(* IEC 61131-3 sources: PLC-IsaVODE/PLC-IsaVODE/samples/plc-programs (part 2) *)

(* ---- 251-SETUP_LANGUAGE.ST ---- *)
TYPE oscat_LANGUAGE:
	STRUCT
		DEFAULT 	: INT;
		LMAX    	: INT;
	END_STRUCT;
END_TYPE

FUNCTION_BLOCK SETUP_LANGUAGE_Block

	VAR_IN_OUT
		LANGUAGE :	oscat_LANGUAGE;
	END_VAR

	VAR
		init :	BOOL;
	END_VAR

	IF init THEN RETURN; END_IF;
	init := TRUE;

	LANGUAGE.DEFAULT  := 1; (* 1=english, 2=german 3=french *)
	LANGUAGE.LMAX := 3;

END_FUNCTION_BLOCK

PROGRAM program0

	VAR
		LANGUAGE :	oscat_LANGUAGE;
		func_block : SETUP_LANGUAGE_Block;
	END_VAR
		func_block.LANGUAGE  := LANGUAGE;
		func_block();
		LANGUAGE := func_block.LANGUAGE;

END_PROGRAM

CONFIGURATION Config0

	RESOURCE Res0 ON PLC
		TASK task0(INTERVAL := T#20ms,PRIORITY := 0);
		PROGRAM instance0 WITH task0 : program0;
	END_RESOURCE

END_CONFIGURATION

(* ---- 253-ENERGY.ST ---- *)
FUNCTION_BLOCK ENERGY
	VAR_INPUT
		J :	REAL;
		C :	REAL;
		WH :	REAL;
	END_VAR

	VAR_OUTPUT
		YJ :	REAL;
		YC :	REAL;
		YWH :	REAL;
	END_VAR

	YJ := J + Wh * 3600.0 + C * 4.1868;
	YC := YJ * 0.238845896627496;
	YWh := YJ * 2.7777777778E-004;
END_FUNCTION_BLOCK

PROGRAM program0
  VAR
		J  :	REAL;
		C  :	REAL;
		WH :	REAL;

		YJ  :	REAL;
		YC  :	REAL;
		YWH :	REAL;
	func_block : ENERGY;
  END_VAR
	func_block.J  :=J ;
	func_block.C  :=C ;
	func_block.WH :=WH;
	func_block();
	YJ  := func_block.YJ ;
	YC  := func_block.YC ;
	YWH := func_block.YWH;

END_PROGRAM

CONFIGURATION Config0
	RESOURCE Res0 ON PLC
		TASK task0(INTERVAL := T#20ms,PRIORITY := 0);
		PROGRAM instance0 WITH task0 : program0;
	END_RESOURCE
END_CONFIGURATION

(* ---- 257-FINDB_NONUM.ST ---- *)
FUNCTION_BLOCK FINDB_NONUM_Block

	VAR_INPUT
		STR :	STRING;
	END_VAR

	VAR_OUTPUT
		FINDB_NONUM :	INT;
	END_VAR

	VAR
		pos :	INT;
		x :	INT;
	END_VAR

	pos := LEN(str);
	WHILE (pos >=1) DO
		x :=GET_CHAR(str,pos);
		IF (X < 48 AND X <> 46) OR X > 57 THEN
			findB_nonum := pos;
			RETURN;
		END_IF;
	pos := pos -1;
	END_WHILE;
	findB_nonum := 0;

END_FUNCTION_BLOCK

PROGRAM program0
	VAR
		STR :	STRING;

		FINDB_NONUM :	INT;

		func_block : FINDB_NONUM_Block;
	END_VAR
	func_block.STR := STR;
	func_block();
	FINDB_NONUM  := func_block.FINDB_NONUM;
END_PROGRAM

CONFIGURATION Config0
	RESOURCE Res0 ON PLC
		TASK task0(INTERVAL := T#20ms,PRIORITY := 0);
		PROGRAM instance0 WITH task0 : program0;
	END_RESOURCE
END_CONFIGURATION

(* ---- 258-HYST_1.ST ---- *)
FUNCTION_BLOCK HYST_1_Block

	VAR_INPUT
		IN :	REAL;
		HIGH :	REAL;
		LOW :	REAL;
	END_VAR

	VAR_OUTPUT
		Q :	BOOL;
		WIN :	BOOL;
	END_VAR

	IF in < low THEN
		Q := FALSE;
		win := FALSE;
	ELSIF in > high THEN
		Q := TRUE;
		win := FALSE;
	ELSE
		win := TRUE;
	END_IF;

END_FUNCTION_BLOCK

PROGRAM program0
	VAR
		IN :	REAL;
		HIGH :	REAL;
		LOW :	REAL;
		Q :	BOOL;
		WIN :	BOOL;
		func_block : HYST_1_Block;
	END_VAR
	func_block.IN := IN;
	func_block.HIGH := HIGH;
	func_block.LOW := LOW;
	func_block();
	Q  := func_block.Q;
	WIN  := func_block.WIN;
END_PROGRAM

CONFIGURATION Config0
	RESOURCE Res0 ON PLC
		TASK task0(INTERVAL := T#20ms,PRIORITY := 0);
		PROGRAM instance0 WITH task0 : program0;
	END_RESOURCE
END_CONFIGURATION

(* ---- 260-V3_SUB.ST ---- *)
TYPE oscat_vector_3:
	STRUCT
		X : REAL;
		Y : REAL;
		Z : REAL;
	END_STRUCT;
END_TYPE

FUNCTION_BLOCK V3_SUB_Block

	VAR_INPUT
		A :	oscat_vector_3;
		B :	oscat_vector_3;
	END_VAR

	VAR_OUTPUT
		V3_SUB :	oscat_vector_3;
	END_VAR

	V3_SUB.X := A.X - B.X;
	V3_SUB.Y := A.Y - B.Y;
	V3_SUB.Z := A.Z - B.Z;

END_FUNCTION_BLOCK

PROGRAM program0
  	VAR
		A :	oscat_vector_3;
		B :	oscat_vector_3;
		V3_SUB :	oscat_vector_3;
		func_block : V3_SUB_Block;
  	END_VAR
	func_block.A := A;
	func_block.B := B;
	func_block();
	V3_SUB := func_block.V3_SUB;
END_PROGRAM

CONFIGURATION Config0
  RESOURCE Res0 ON PLC
    TASK task0(INTERVAL := T#20ms,PRIORITY := 0);
    PROGRAM instance0 WITH task0 : program0;
  END_RESOURCE
END_CONFIGURATION

(* ---- 261-A_TRIG.ST ---- *)
FUNCTION_BLOCK A_TRIG

	VAR_INPUT
		IN :	REAL;
		RES :	REAL;
	END_VAR

	VAR_OUTPUT
		Q :	BOOL;
		D :	REAL;
	END_VAR

	VAR
		last_in :	REAL;
	END_VAR

	D := IN - LAST_IN;
	IF ABS(D) >= res THEN
		Q := TRUE;
		last_in := IN;
	ELSE
		Q := FALSE;
	END_IF;

END_FUNCTION_BLOCK

PROGRAM program0
	VAR
	    LocalVar0 : REAL;
		LocalVar1 : REAL;
		LocalOUT1  : BOOL;
		LocalOUT2  : REAL;
		func_block : A_TRIG;
  	END_VAR
	func_block.IN := LocalVar0;
    func_block.RES := LocalVar1;
	func_block();
	LocalOUT1 := func_block.Q;
	LocalOUT2 := func_block.D;
END_PROGRAM

CONFIGURATION Config0
  	RESOURCE Res0 ON PLC
    	TASK task0(INTERVAL := T#20ms,PRIORITY := 0);
    	PROGRAM instance0 WITH task0 : program0;
  	END_RESOURCE
END_CONFIGURATION

(* ---- 265-INTERLOCK.ST ---- *)
FUNCTION_BLOCK INTERLOCK_Block

	VAR_INPUT
		I1 :	BOOL;
		I2 :	BOOL;
		TL :	TIME;
	END_VAR

	VAR_OUTPUT
		Q1 :	BOOL;
		Q2 :	BOOL;
	END_VAR

	VAR
		T1 :	TOF;
		T2 :	TOF;
	END_VAR

	T1(IN := I1, PT := TL);
	T2(IN := I2, PT := TL);

	Q1 := I1 AND NOT t2.Q;
	Q2 := I2 AND NOT t1.Q;

END_FUNCTION_BLOCK

PROGRAM program0
	VAR
		I1 :	BOOL;
		I2 :	BOOL;
		TL :	TIME;
		Q1 :	BOOL;
		Q2 :	BOOL;
		func_block : INTERLOCK_Block;
  	END_VAR
	func_block.I1  :=I1;
	func_block.I2  :=I2;
	func_block.TL  :=TL;
	func_block();
	Q1 := func_block.Q1;
	Q2 := func_block.Q2;
END_PROGRAM

CONFIGURATION Config0
	RESOURCE Res0 ON PLC
		TASK task0(INTERVAL := T#20ms,PRIORITY := 0);
		PROGRAM instance0 WITH task0 : program0;
	END_RESOURCE
END_CONFIGURATION

(* ---- 266-CMUL.ST ---- *)
TYPE oscat_complex :
  STRUCT
	re : REAL;
	im : REAL;
  END_STRUCT;
END_TYPE

FUNCTION_BLOCK CMUL_Block

	VAR_INPUT
		X :	oscat_complex;
		Y :	oscat_complex;
	END_VAR

	VAR_OUTPUT
		CMUL :	oscat_complex;
	END_VAR

	CMUL.re := X.re * Y.re - X.im * Y.im;
	CMUL.im := X.re * Y.im + X.im * Y.re;
END_FUNCTION_BLOCK

PROGRAM program0
  VAR
    LocalVar0 : oscat_complex;
	LocalVar1 : oscat_complex;
	LocalOUT  : oscat_complex;
	func_block : CMUL_Block;
  END_VAR
	func_block.X  := LocalVar0;
	func_block.Y  := LocalVar1;
	func_block();
	LocalOUT := func_block.CMUL;
END_PROGRAM

CONFIGURATION Config0
  RESOURCE Res0 ON PLC
    TASK task0(INTERVAL := T#20ms,PRIORITY := 0);
    PROGRAM instance0 WITH task0 : program0;
  END_RESOURCE
END_CONFIGURATION

(* ---- 268-IS_UPPER.ST ---- *)
FUNCTION SETUP_EXTENDED_ASCII:BOOL

	VAR_INPUT
		X :	BOOL;
	END_VAR

	SETUP_EXTENDED_ASCII := X OR TRUE;

END_FUNCTION

FUNCTION ISC_UPPER:BOOL

	VAR_INPUT
		IN :	BYTE;
	END_VAR

	IF SETUP_EXTENDED_ASCII(FALSE) THEN
		ISC_UPPER :=  ((in > BYTE#64) AND (in < BYTE#91)) OR (((in > BYTE#191) AND (in < BYTE#223)) AND (in <> BYTE#215));
	ELSE
		ISC_UPPER := ((in > BYTE#64) AND (in < BYTE#91));
	END_IF;

END_FUNCTION

FUNCTION_BLOCK IS_UPPER

	VAR_INPUT
		STR :	STRING;
	END_VAR

	VAR_OUTPUT
		IS_UPPER :	BOOL;
	END_VAR

	VAR
		pos :	INT;
		I :	INT;
	END_VAR

	I := LEN(str);
	FOR pos := 1 TO I DO
		IF NOT ISC_UPPER(INT_TO_BYTE(GET_CHAR(str,pos))) THEN
			IS_UPPER := FALSE;
			RETURN;
		END_IF;
	END_FOR;
	IS_UPPER := I>0;

END_FUNCTION_BLOCK

(* ---- 269-IS_CC.ST ---- *)
FUNCTION_BLOCK IS_CC_Block

	VAR_INPUT
		STR :	STRING;
		CMP :	STRING;
	END_VAR

	VAR_OUTPUT
		IS_CC :	BOOL;
	END_VAR

	VAR
		L :	INT;
		pos :	INT;
		temp :	STRING;
	END_VAR

	L := LEN(str);
	FOR pos := 1 TO L DO
		temp := MID(str,1,pos);
		IF FIND(CMP,temp) = 0 THEN
			IS_CC := FALSE;
			RETURN;
		END_IF;
	END_FOR;
	IS_CC := L > 0;

END_FUNCTION_BLOCK

PROGRAM program0

	VAR
		STR :	STRING;
		CMP :	STRING;

		IS_CC :	BOOL;

		func_block : IS_CC_Block;
	END_VAR
	func_block.STR := STR;
	func_block.CMP := CMP;
	func_block();
	IS_CC := func_block.IS_CC;

END_PROGRAM

CONFIGURATION Config0

	RESOURCE Res0 ON PLC
		TASK task0(INTERVAL := T#20ms,PRIORITY := 0);
		PROGRAM instance0 WITH task0 : program0;
	END_RESOURCE

END_CONFIGURATION

(* ---- 271-IS_NCC.ST ---- *)
FUNCTION_BLOCK IS_NCC_Block

	VAR_INPUT
		STR :	STRING;
		CMP :	STRING;
	END_VAR

	VAR_OUTPUT
		IS_NCC :	BOOL;
	END_VAR

	VAR
		L :	INT;
		pos :	INT;
		temp :	STRING;
	END_VAR

	L := LEN(str);
	FOR pos := 1 TO L DO
		temp := MID(str,1,pos);
		IF FIND(CMP,temp) > 0 THEN
			IS_NCC := FALSE;
			RETURN;
		END_IF;
	END_FOR;
	IS_NCC := TRUE;

END_FUNCTION_BLOCK

PROGRAM program0

	VAR
		STR :	STRING;
		CMP :	STRING;
		IS_NCC :	BOOL;
		func_block : IS_NCC_Block;
	END_VAR
	func_block.STR := STR;
	func_block.CMP := CMP;
	func_block();
	IS_NCC := func_block.IS_NCC;

END_PROGRAM

CONFIGURATION Config0

	RESOURCE Res0 ON PLC
		TASK task0(INTERVAL := T#20ms,PRIORITY := 0);
		PROGRAM instance0 WITH task0 : program0;
	END_RESOURCE

END_CONFIGURATION

(* ---- 273-TONOF.ST ---- *)
FUNCTION_BLOCK TONOF

	VAR_INPUT
		IN :	BOOL;
		T_ON :	TIME;
		T_OFF :	TIME;
	END_VAR

	VAR_OUTPUT
		Q :	BOOL;
	END_VAR

	VAR
		X :	TON;
		old :	BOOL;
		mode :	BOOL;
	END_VAR

	IF IN XOR old THEN
	X(IN := FALSE, PT := SEL_TIME(IN,T_OFF,T_ON));
	mode := IN;
	old := IN;
	END_IF;
	X(IN := TRUE);
	IF X.Q THEN Q := mode;END_IF;

END_FUNCTION_BLOCK

PROGRAM program0
  VAR
	IN :	BOOL;
	T_ON :	TIME;
	T_OFF :	TIME;
	Q :	BOOL;
	func_block : TONOF;
  END_VAR
	func_block.IN  :=IN ;
	func_block.T_ON  :=T_ON ;
	func_block.T_OFF  :=T_OFF ;
	func_block();
	Q := func_block.Q;

END_PROGRAM

CONFIGURATION Config0
	RESOURCE Res0 ON PLC
		TASK task0(INTERVAL := T#20ms,PRIORITY := 0);
		PROGRAM instance0 WITH task0 : program0;
	END_RESOURCE
END_CONFIGURATION

(* ---- 278-DWORD_TO_STRB.ST ---- *)
FUNCTION_BLOCK DWORD_TO_STRB_Block
	VAR_INPUT
		IN :	DWORD;
	END_VAR

	VAR_OUTPUT
		DWORD_TO_STRB :	STRING;
	END_VAR

	VAR
		i :	INT;
	END_VAR

	DWORD_TO_STRB :='';
	FOR i := 1 TO 32 DO
		IF (in AND DWORD#16#8000_0000) > DWORD#0 THEN
			DWORD_TO_STRB := CONCAT(DWORD_TO_STRB,'1');
		ELSE
			DWORD_TO_STRB := CONCAT(DWORD_TO_STRB,'0');
		END_IF;
		in := SHL(in, 1);
	END_FOR;
END_FUNCTION_BLOCK

PROGRAM program0
  VAR
    IN :	DWORD;

	DWORD_TO_STRB :	STRING;
	func_block : DWORD_TO_STRB_Block;
  END_VAR
	func_block.IN  := IN;
	func_block();
	DWORD_TO_STRB := func_block.DWORD_TO_STRB;
END_PROGRAM

CONFIGURATION Config0
  RESOURCE Res0 ON PLC
    TASK task0(INTERVAL := T#20ms,PRIORITY := 0);
    PROGRAM instance0 WITH task0 : program0;
  END_RESOURCE
END_CONFIGURATION

(* ---- 279-STAIR2.ST ---- *)
FUNCTION FLOOR : INT
	VAR_INPUT
		x : REAL;
	END_VAR

	FLOOR := REAL_TO_INT(X);
	IF INT_TO_REAL(FLOOR) > X THEN
		floor := floor - 1;
	END_IF;
END_FUNCTION

FUNCTION_BLOCK STAIR2_Block

	VAR_INPUT
		X :	REAL;
		D :	REAL;
	END_VAR

	VAR_OUTPUT
		Y :	REAL;
	END_VAR

	IF D > 0.0 THEN
		IF X >= Y + D OR X <= Y - D THEN Y := INT_TO_REAL(FLOOR(X/D)) * D; END_IF;
	ELSE
		Y := X;
	END_IF;

END_FUNCTION_BLOCK

PROGRAM program0

	VAR
		X :	REAL;
		D :	REAL;
		Y :	REAL;
		func_block : STAIR2_Block;
	END_VAR
	func_block.X := X;
	func_block.D := D;
	func_block();
	Y := func_block.Y;

END_PROGRAM

CONFIGURATION Config0

	RESOURCE Res0 ON PLC
		TASK task0(INTERVAL := T#20ms,PRIORITY := 0);
		PROGRAM instance0 WITH task0 : program0;
	END_RESOURCE

END_CONFIGURATION

(* ---- 280-DEC_TO_BYTE.ST ---- *)
FUNCTION_BLOCK DEC_TO_BYTE_Block
	VAR_INPUT
		DEC :	STRING;
	END_VAR

	VAR_OUTPUT
		DEC_TO_BYTE :	BYTE;
	END_VAR

	VAR
		i :	INT;
		X :	INT;
		stop :	INT;
	END_VAR

	DEC_TO_BYTE := BYTE#0;
	stop := LEN(DEC);
	FOR I := 1 TO stop DO
		X := GET_CHAR(DEC,I);
		IF X > 47 AND X < 58 THEN
			DEC_TO_BYTE := INT_TO_BYTE(_BYTE_TO_INT(DEC_TO_BYTE) * 10 + X - 48);
		END_IF;
	END_FOR;

END_FUNCTION_BLOCK

PROGRAM program0
  VAR
    LocalVar0 : STRING;
	LocalOUT  : BYTE;
	func_block : DEC_TO_BYTE_Block;
  END_VAR
	func_block.DEC  := LocalVar0;
	func_block();
	LocalOUT := func_block.DEC_TO_BYTE;
END_PROGRAM

CONFIGURATION Config0
  RESOURCE Res0 ON PLC
    TASK task0(INTERVAL := T#20ms,PRIORITY := 0);
    PROGRAM instance0 WITH task0 : program0;
  END_RESOURCE
END_CONFIGURATION

(* ---- 281-BYTE_TO_STRB.ST ---- *)
FUNCTION_BLOCK BYTE_TO_STRB_Block
	VAR_INPUT
		IN :	BYTE;
	END_VAR

	VAR_OUTPUT
		BYTE_TO_STRB :	STRING;
	END_VAR

	VAR
		i :	INT;
	END_VAR

	BYTE_TO_STRB := '';
	FOR i := 1 TO 8 DO
		IF (in AND BYTE#2#1000_0000) = BYTE#2#1000_0000 THEN
			BYTE_TO_STRB := CONCAT(BYTE_TO_STRB,'1');
		ELSE
			BYTE_TO_STRB := CONCAT(BYTE_TO_STRB,'0');
		END_IF;
		in := SHL(in, 1);
	END_FOR;

END_FUNCTION_BLOCK

PROGRAM program0
  VAR
    LocalVar0 : BYTE;
	LocalOUT  : STRING;
	func_block : BYTE_TO_STRB_Block;
  END_VAR
	func_block.IN  := LocalVar0;
	func_block();
	LocalOUT := func_block.BYTE_TO_STRB;

END_PROGRAM

CONFIGURATION Config0
  RESOURCE Res0 ON PLC
    TASK task0(INTERVAL := T#20ms,PRIORITY := 0);
    PROGRAM instance0 WITH task0 : program0;
  END_RESOURCE
END_CONFIGURATION

(* ---- 282-SW_RECONFIG.ST ---- *)
FUNCTION_BLOCK SW_RECONFIG_Block

	VAR_INPUT
		IN :	BOOL;
		TD :	TIME;
		TR :	TIME;
	END_VAR

	VAR_OUTPUT
		Q :	BOOL;
	END_VAR

	VAR
		T1 :	TON;
		T2 :	TON;
		INV :	BOOL;
	END_VAR

	t1(in := IN, PT := TD);

	IF tr > t#0s THEN
		Q := t1.Q XOR inv;
		T2(in := Q, pt := TR);
		IF T2.Q THEN INV := NOT INV; END_IF;
	ELSE
		Q := t1.Q;
	END_IF;

END_FUNCTION_BLOCK

PROGRAM program0
	VAR
		IN :	BOOL;
		TD :	TIME;
		TR :	TIME;
		Q :	BOOL;

		func_block : SW_RECONFIG_Block;
	END_VAR
	func_block.IN := IN;
	func_block.TD := TD;
	func_block.TR := TR ;

	func_block();
	Q  := func_block.Q;

END_PROGRAM

CONFIGURATION Config0
	RESOURCE Res0 ON PLC
		TASK task0(INTERVAL := T#20ms,PRIORITY := 0);
		PROGRAM instance0 WITH task0 : program0;
	END_RESOURCE
END_CONFIGURATION

(* ---- 283-CINV.ST ---- *)
TYPE oscat_complex :
  STRUCT
	re : REAL;
	im : REAL;
  END_STRUCT;
END_TYPE

FUNCTION_BLOCK CINV_Block

	VAR_INPUT
		X :	oscat_complex;
	END_VAR

	VAR_OUTPUT
		CINV :	oscat_complex;
	END_VAR

	VAR
		temp :	REAL;
	END_VAR

	temp := X.re * X.re + X.im * X.im;
	IF temp = 0.0 THEN CINV.re := 0.0;CINV.im := 0.0;RETURN;END_IF;
	CINV.re := X.re / temp;
	CINV.im := -X.im / temp;

END_FUNCTION_BLOCK

PROGRAM program0
  VAR
    LocalVar0 : oscat_complex;
	LocalOUT  : oscat_complex;
	func_block : CINV_Block;
  END_VAR
	func_block.X  := LocalVar0;
	func_block();
	LocalOUT := func_block.CINV;
END_PROGRAM

CONFIGURATION Config0
  RESOURCE Res0 ON PLC
    TASK task0(INTERVAL := T#20ms,PRIORITY := 0);
    PROGRAM instance0 WITH task0 : program0;
  END_RESOURCE
END_CONFIGURATION

(* ---- 284-V3_XPRO.ST ---- *)
TYPE oscat_vector_3 :
	STRUCT
		X : REAL;
		Y : REAL;
		Z : REAL;
	END_STRUCT;
END_TYPE

FUNCTION_BLOCK V3_XPRO_Block
	VAR_INPUT
		A :	oscat_vector_3;
		B :	oscat_vector_3;
	END_VAR

	VAR_OUTPUT
		V3_XPRO :	oscat_vector_3;
	END_VAR

	V3_XPRO.X := A.Y * B.Z - A.Z * B.Y;
	V3_XPRO.Y := A.Z * B.X - A.X * B.Z;
	V3_XPRO.Z := A.X * B.Y - A.Y * B.X;

END_FUNCTION_BLOCK

PROGRAM program0
  	VAR
		A :	oscat_vector_3;
		B :	oscat_vector_3;
		V3_XPRO :	oscat_vector_3;
		func_block : V3_XPRO_Block;
  	END_VAR
	func_block.A := A;
	func_block.B := B;
	func_block();
	V3_XPRO := func_block.V3_XPRO;
END_PROGRAM

CONFIGURATION Config0
  RESOURCE Res0 ON PLC
    TASK task0(INTERVAL := T#20ms,PRIORITY := 0);
    PROGRAM instance0 WITH task0 : program0;
  END_RESOURCE
END_CONFIGURATION

(* ---- 288-DEC_4.ST ---- *)
FUNCTION_BLOCK DEC_4
	VAR_INPUT
		D :	BOOL;
		A0 :	BOOL;
		A1 :	BOOL;
	END_VAR

	VAR_OUTPUT
		Q0 :	BOOL;
		Q1 :	BOOL;
		Q2 :	BOOL;
		Q3 :	BOOL;
	END_VAR

	Q0 := D AND NOT A0 AND NOT A1;
	Q1 := D AND A0 AND NOT A1;
	Q2 := D AND NOT A0 AND A1;
	Q3 := D AND A0 AND A1;
END_FUNCTION_BLOCK

PROGRAM program0
  VAR
	D :	BOOL;
	A0 :	BOOL;
	A1 :	BOOL;

	Q0 :	BOOL;
	Q1 :	BOOL;
	Q2 :	BOOL;
	Q3 :	BOOL;

	func_block : DEC_4;
  END_VAR
	func_block.D   := D  ;
	func_block.A0  := A0  ;
	func_block.A1  := A1  ;
	func_block();
	Q0:= func_block.Q0;
	Q1:= func_block.Q1;
	Q2:= func_block.Q2;
	Q3:= func_block.Q3;
END_PROGRAM

CONFIGURATION Config0
  RESOURCE Res0 ON PLC
    TASK task0(INTERVAL := T#20ms,PRIORITY := 0);
    PROGRAM instance0 WITH task0 : program0;
  END_RESOURCE
END_CONFIGURATION

(* ---- 291-FF_D2E.ST ---- *)
FUNCTION_BLOCK FF_D2E
	VAR_INPUT
		D0 :	BOOL;
		D1 :	BOOL;
		CLK :	BOOL;
		RST :	BOOL;
	END_VAR

	VAR_OUTPUT
		Q0 :	BOOL;
		Q1 :	BOOL;
	END_VAR

	VAR
		edge :	BOOL;
	END_VAR

	IF rst THEN
		Q0 := FALSE;
		Q1 := FALSE;
	ELSIF clk AND NOT edge THEN
		Q0 := D0;
		Q1 := D1;
	END_IF;
	edge := CLK;

END_FUNCTION_BLOCK

PROGRAM program0
  VAR
	D0  :	BOOL;
	D1  :	BOOL;
	CLK :	BOOL;
	RST :	BOOL;

	Q0 :	BOOL;
	Q1 :	BOOL;

	func_block : FF_D2E;
  END_VAR
	func_block.D0  :=D0 ;
	func_block.D1  :=D1 ;
	func_block.CLK :=CLK;
	func_block.RST :=RST;
	func_block();
	Q0 := func_block.Q0;
	Q1 := func_block.Q1;
END_PROGRAM

CONFIGURATION Config0
  RESOURCE Res0 ON PLC
    TASK task0(INTERVAL := T#20ms,PRIORITY := 0);
    PROGRAM instance0 WITH task0 : program0;
  END_RESOURCE
END_CONFIGURATION

(* ---- 292-HYST_2.ST ---- *)
FUNCTION_BLOCK HYST_2_Block

	VAR_INPUT
		IN :	REAL;
		VAL :	REAL;
		HYS :	REAL;
	END_VAR

	VAR_OUTPUT
		Q :	BOOL;
		WIN :	BOOL;
	END_VAR

	VAR
		tmp :	REAL;
	END_VAR

	tmp := val - hys * 0.5;
	IF in < tmp THEN
		Q := FALSE;
		win := FALSE;
	ELSIF in > tmp + hys THEN
		Q := TRUE;
		win := FALSE;
	ELSE
		win := TRUE;
	END_IF;

END_FUNCTION_BLOCK

PROGRAM program0
	VAR
		IN :	REAL;
		VAL :	REAL;
		HYS :	REAL;
		Q :	BOOL;
		WIN :	BOOL;
		func_block : HYST_2_Block;
	END_VAR
	func_block.IN := IN;
	func_block.VAL := VAL;
	func_block.HYS := HYS;
	func_block();
	Q  := func_block.Q;
	WIN  := func_block.WIN;
END_PROGRAM

CONFIGURATION Config0
	RESOURCE Res0 ON PLC
		TASK task0(INTERVAL := T#20ms,PRIORITY := 0);
		PROGRAM instance0 WITH task0 : program0;
	END_RESOURCE
END_CONFIGURATION

(* ---- 294-FF_RSE.ST ---- *)
FUNCTION_BLOCK FF_RSE
	VAR_INPUT
		CS :	BOOL;
		CR :	BOOL;
		RST :	BOOL;
	END_VAR

	VAR_OUTPUT
		Q :	BOOL;
	END_VAR

	VAR
		es :	BOOL;
		er :	BOOL;
	END_VAR

	IF rst THEN
		(* asynchronous reset *)
		Q := FALSE;
	ELSIF CR AND NOT er THEN
		(* rising edge on CR *)
		Q := FALSE;
	ELSIF CS AND NOT es THEN
		(* rising edge on CS *)
		Q := TRUE;
	END_IF;

	es := CS;
	er := CR;
END_FUNCTION_BLOCK

PROGRAM program0
  VAR
	CS  :	BOOL;
	CR  :	BOOL;
	RST :	BOOL;

	Q :	BOOL;

	func_block : FF_RSE;
  END_VAR
	func_block.CS  :=CS ;
	func_block.CR  :=CR ;
	func_block.RST :=RST;
	func_block();
	Q := func_block.Q;
END_PROGRAM

CONFIGURATION Config0
  RESOURCE Res0 ON PLC
    TASK task0(INTERVAL := T#20ms,PRIORITY := 0);
    PROGRAM instance0 WITH task0 : program0;
  END_RESOURCE
END_CONFIGURATION

(* ---- 296-BUFFER_CLEAR_NW.ST ---- *)
TYPE
  oscat_NW_BUF_LONG  : ARRAY [0..4095] OF BYTE;
END_TYPE

FUNCTION_BLOCK _BUFFER_CLEAR_NW
	VAR_INPUT
		SIZE :	UINT;
	END_VAR

	VAR_OUTPUT
		BUFFER_CLEAR :	BOOL;
	END_VAR

	VAR_IN_OUT
		PT :	oscat_NW_BUF_LONG;
	END_VAR

	VAR
		err :	INT;
		result :	WORD;
	END_VAR
	result:=MEMSET(err,BYTE#00,UINT_TO_DINT(size),pt[0]);
	BUFFER_CLEAR := (err = 0);
END_FUNCTION_BLOCK

PROGRAM program0
  VAR
	SIZE :	UINT;

	BUFFER_CLEAR :	BOOL;

	PT :	oscat_NW_BUF_LONG;

	func_block : _BUFFER_CLEAR_NW;
  END_VAR
	func_block.SIZE  :=SIZE ;
	func_block.PT  :=PT ;
	func_block();
	PT := func_block.PT;
	BUFFER_CLEAR := func_block.BUFFER_CLEAR;
END_PROGRAM

CONFIGURATION Config0
  RESOURCE Res0 ON PLC
    TASK task0(INTERVAL := T#20ms,PRIORITY := 0);
    PROGRAM instance0 WITH task0 : program0;
  END_RESOURCE
END_CONFIGURATION

(* ---- 298-FF_JKE.ST ---- *)
FUNCTION_BLOCK FF_JKE
	VAR_INPUT
		SET :	BOOL;
		J :	BOOL;
		CLK :	BOOL;
		K :	BOOL;
		RST :	BOOL;
	END_VAR

	VAR_OUTPUT
		Q :	BOOL;
	END_VAR

	VAR
		edge :	BOOL;
	END_VAR

	IF rst OR set THEN
		Q := NOT rst;
	ELSIF clk AND NOT edge THEN
		IF J XOR K THEN Q := J;
		ELSE Q := K XOR Q;
		END_IF;
	END_IF;
	edge := CLK;

END_FUNCTION_BLOCK

PROGRAM program0
  VAR
		SET :	BOOL;
		J   :	BOOL;
		CLK :	BOOL;
		K   :	BOOL;
		RST :	BOOL;

		Q :	BOOL;

	func_block : FF_JKE;
  END_VAR
	func_block.SET :=SET;
	func_block.J   :=J  ;
	func_block.CLK :=CLK;
	func_block.K   :=K  ;
	func_block.RST :=RST;
	func_block();
	Q := func_block.Q;
END_PROGRAM

CONFIGURATION Config0
  RESOURCE Res0 ON PLC
    TASK task0(INTERVAL := T#20ms,PRIORITY := 0);
    PROGRAM instance0 WITH task0 : program0;
  END_RESOURCE
END_CONFIGURATION

(* ---- 299-OCT_TO_DWORD.ST ---- *)
FUNCTION_BLOCK OCT_TO_DWORD_Block

	VAR_INPUT
		OCT :	STRING;
	END_VAR

	VAR_OUTPUT
		OCT_TO_DWORD :	DWORD;
	END_VAR

	VAR
		i :	INT;
		stop :	INT;
		X :	INT;
	END_VAR

	OCT_TO_DWORD := DWORD#0;
	stop := LEN(oct);
	FOR I := 1 TO stop DO
		X := GET_CHAR(oct,I);
		(* calculate the value of the digit *)
		IF X > 47 AND x < 56 THEN
			OCT_TO_DWORD := SHL_DWORD(OCT_TO_DWORD,3) OR INT_TO_DWORD(X - 48);
		END_IF;
	END_FOR;

END_FUNCTION_BLOCK

PROGRAM program0
  VAR
    OCT : STRING;
    OCT_TO_DWORD : DWORD;
	func_block : OCT_TO_DWORD_Block;
  END_VAR

  	func_block.OCT := '125';
	func_block();
	OCT_TO_DWORD := func_block.OCT_TO_DWORD;
END_PROGRAM

CONFIGURATION Config0
	RESOURCE Res0 ON PLC
		TASK task0(INTERVAL := T#20ms,PRIORITY := 0);
		PROGRAM instance0 WITH task0 : program0;
	END_RESOURCE
END_CONFIGURATION

(* ---- 3-IS_LOWER.ST ---- *)
FUNCTION_BLOCK IS_LOWER

VAR_INPUT
	STR :	STRING;
END_VAR

VAR_OUTPUT
	IS_LOWER :	BOOL;
END_VAR

VAR
	pos :	INT;
	I :	INT;
END_VAR

I := LEN(str);
FOR pos := 1 TO I DO
	IF NOT ISC_LOWER(INT_TO_BYTE(GET_CHAR(str,pos))) THEN
		IS_LOWER := FALSE;
		RETURN;
	END_IF;
END_FOR;
IS_LOWER := I>0;

END_FUNCTION_BLOCK

(* ---- 302-MD5_TO_STRH.ST ---- *)
FUNCTION_BLOCK MD5_TO_STRH

	VAR_INPUT
		MD5 :	oscat_aB0_15;
	END_VAR

	VAR_OUTPUT
		MD5_TO_STRH :	oscat_STRING32;
	END_VAR

	VAR
		buf :	oscat_aB0_31;
		x :	INT;
		BUF_TO_STRING :	BUF_TO_STRING;
		i :	INT;
		tmp :	INT;
	END_VAR

	x := 0;
	FOR i := 0 TO 15 DO;
		tmp := BYTE_TO_INT(SHR_BYTE(MD5[i],4));
		buf[x] := INT_TO_BYTE(tmp + SEL(tmp <= 9,87,48));
		x := x + 1;
		tmp := BYTE_TO_INT(MD5[i] AND BYTE#2#1111);
		buf[x] := INT_TO_BYTE(tmp + SEL(tmp <= 9,87,48));
		x := x + 1;
	END_FOR;

	FOR x := 0 TO 1 DO
		BUF_TO_STRING.REQ := x > 0;
		BUF_TO_STRING.BUF_FORMAT := TRUE;
		BUF_TO_STRING.BUF_OFFS := DINT#0;
		BUF_TO_STRING.BUF_CNT := DINT#32;
		BUF_TO_STRING.BUFFER := buf;
		BUF_TO_STRING.DST := MD5_TO_STRH;
		BUF_TO_STRING();
		buf := BUF_TO_STRING.BUFFER;
		MD5_TO_STRH := BUF_TO_STRING.DST;
	END_FOR;

END_FUNCTION_BLOCK

(* ---- 303-FINDB.ST ---- *)
FUNCTION_BLOCK FINDB_Block

	VAR_INPUT
		STR1 :	STRING;
		STR2 :	STRING;
	END_VAR

	VAR_OUTPUT
		FINDB :	INT;
	END_VAR

	VAR
		pos :	INT;
		length :	INT;
		string_temp :	STRING;
	END_VAR

	length := LEN(str2);
	pos := LEN(str1) - length +1;
	WHILE (pos >= 1) DO
		string_temp := MID(str1,length,pos);
		IF EQ_STRING(string_temp,str2) THEN
			FindB := pos;
			RETURN;
		END_IF;
	pos := pos -1;
	END_WHILE;
	FindB := 0;

END_FUNCTION_BLOCK

PROGRAM program0
  VAR
		STR1 :	STRING;
		STR2 :	STRING;

		FINDB :	INT;

	func_block : FINDB_Block;
  END_VAR
	func_block.STR1  := STR1;
	func_block.STR2  := STR2;
	func_block();
	FINDB := func_block.FINDB;
END_PROGRAM

CONFIGURATION Config0

	RESOURCE Res0 ON PLC
		TASK task0(INTERVAL := T#20ms,PRIORITY := 0);
		PROGRAM instance0 WITH task0 : program0;
	END_RESOURCE
END_CONFIGURATION

(* ---- 305-SEL2_OF_3B.ST ---- *)
FUNCTION_BLOCK SEL2_OF_3B_Block

	VAR_INPUT
		IN1 :	BOOL;
		IN2 :	BOOL;
		IN3 :	BOOL;
		TD :	TIME;
	END_VAR

	VAR_OUTPUT
		Q :	BOOL;
		W :	BOOL;
	END_VAR

	VAR
		TDEL :	TON;
	END_VAR

	Q := (IN1 AND IN2) OR (IN1 AND IN3) OR (IN2 AND IN3);
	TDEL(IN := (in1 XOR in2) OR (in1 XOR in3) OR (in2 XOR in3), PT := TD);
	W := TDEL.Q;

END_FUNCTION_BLOCK

PROGRAM program0

	VAR
		IN1 :	BOOL;
		IN2 :	BOOL;
		IN3 :	BOOL;
		TD :	TIME;
		Q :	BOOL;
		W :	BOOL;
		func_block : SEL2_OF_3B_Block;
  	END_VAR
	func_block.IN1  :=IN1;
	func_block.IN2  :=IN2;
	func_block.IN3  :=IN3;
	func_block.TD  :=TD;
	func_block();
	Q := func_block.Q;
	W := func_block.W;

END_PROGRAM

CONFIGURATION Config0

	RESOURCE Res0 ON PLC
		TASK task0(INTERVAL := T#20ms,PRIORITY := 0);
		PROGRAM instance0 WITH task0 : program0;
	END_RESOURCE

END_CONFIGURATION

(* ---- 306-ARRAY_SUM.ST ---- *)
TYPE
	oscat_pt_ARRAY: ARRAY [1..100] OF REAL;
END_TYPE

FUNCTION_BLOCK ARRAY_SUM_Block
	VAR_IN_OUT
		PT :	oscat_pt_ARRAY;
	END_VAR

	VAR_INPUT
		SIZE :	UINT;
	END_VAR

	VAR_OUTPUT
		ARRAY_SUM :	REAL;
	END_VAR

	VAR
		i :	INT;
		stop :	INT;
	END_VAR

	stop :=LIMIT_INT(1,UINT_TO_INT(size),1000);

	array_sum := pt[1];
	FOR i := 2 TO stop DO
		array_sum := array_sum + pt[i];
	END_FOR;
END_FUNCTION_BLOCK

PROGRAM program0
  VAR
    LocalVar0 : oscat_pt_ARRAY;
    LocalVar1 : UINT;
	LocalOUT  : REAL;
	func_block : ARRAY_SUM_Block;
  END_VAR
	func_block.pt := LocalVar0;
	func_block.size := LocalVar1;
	func_block();
	LocalOUT := func_block.ARRAY_SUM;

END_PROGRAM

CONFIGURATION Config0
  RESOURCE Res0 ON PLC
    TASK task0(INTERVAL := T#20ms,PRIORITY := 0);
    PROGRAM instance0 WITH task0 : program0;
  END_RESOURCE
END_CONFIGURATION

(* ---- 307-ARRAY_MAX.ST ---- *)
TYPE
	oscat_pt_ARRAY: ARRAY [1..100] OF REAL;
END_TYPE

FUNCTION_BLOCK ARRAY_MAX_Block
	VAR_IN_OUT
		PT :	oscat_pt_ARRAY;
	END_VAR

	VAR_INPUT
		SIZE :	UINT;
	END_VAR

	VAR_OUTPUT
		ARRAY_MAX :	REAL;
	END_VAR

	VAR
		i :	INT;
		stop :	INT;
	END_VAR

	stop :=LIMIT_INT(1,UINT_TO_INT(size),1000);

	FOR i := 1 TO stop DO
		IF pt[i] > array_max THEN array_max := pt[i]; END_IF;
	END_FOR;

END_FUNCTION_BLOCK

PROGRAM program0
  VAR
    LocalVar0 : oscat_pt_ARRAY;
    LocalVar1 : UINT;
	LocalOUT  : REAL;
	func_block : ARRAY_MAX_Block;
  END_VAR
	func_block.pt := LocalVar0;
	func_block.size := LocalVar1;
	func_block();
	LocalOUT := func_block.ARRAY_MAX;

END_PROGRAM

CONFIGURATION Config0
  RESOURCE Res0 ON PLC
    TASK task0(INTERVAL := T#20ms,PRIORITY := 0);
    PROGRAM instance0 WITH task0 : program0;
  END_RESOURCE
END_CONFIGURATION

(* ---- 308-DWORD_TO_STRF.ST ---- *)
FUNCTION_BLOCK DWORD_TO_STRF_Block

	VAR_INPUT
		IN :	DWORD;
		N :	INT;
	END_VAR

	VAR_OUTPUT
		DWORD_TO_STRF :	STRING;
	END_VAR

	VAR
		temp :	STRING;
		temp2 :	STRING;
		L : INT;
	END_VAR

	temp := DWORD_TO_STRING(in);
	L := LEN(temp);
	IF N < L THEN
		temp :=RIGHT(temp,N);
		L := N;
	END_IF;

	WHILE L < N DO
		temp2 := temp;
		temp := CONCAT('0', temp2);
		L := L + 1;
	END_WHILE;
	DWORD_TO_STRF := temp;

END_FUNCTION_BLOCK

PROGRAM program0
  VAR
    IN :	DWORD;
	N :		INT;
	DWORD_TO_STRF :	STRING;
	func_block : DWORD_TO_STRF_Block;
  END_VAR
	func_block.IN  := IN;
	func_block.N  := N;
	func_block();
	DWORD_TO_STRF := func_block.DWORD_TO_STRF;
END_PROGRAM

CONFIGURATION Config0
  RESOURCE Res0 ON PLC
    TASK task0(INTERVAL := T#20ms,PRIORITY := 0);
    PROGRAM instance0 WITH task0 : program0;
  END_RESOURCE
END_CONFIGURATION

(* ---- 309-SHA1_TO_STRH.ST ---- *)
FUNCTION_BLOCK SHA1_TO_STRH_Block

	VAR_INPUT
		SHA1 :	oscat_aB0_19;
	END_VAR

	VAR_OUTPUT
		SHA1_TO_STRH :	oscat_STRING40;
	END_VAR

	VAR
		buf :	oscat_aB0_39;
		i :	INT;
		tmp :	INT;
		x :	INT;
		BUF_TO_STRING :	BUF_TO_STRING;
	END_VAR

	x := 0;
	FOR i := 0 TO 19 DO;
		tmp := BYTE_TO_INT(SHR_BYTE(SHA1[i],4));
		buf[x] := INT_TO_BYTE(tmp + SEL(tmp <= 9,87,48));
		x := x + 1;
		tmp := BYTE_TO_INT(SHA1[i] AND BYTE#2#1111);
		buf[x] := INT_TO_BYTE(tmp + SEL(tmp <= 9,87,48));
		x := x + 1;
	END_FOR;

	FOR x := 0 TO 1 DO
		BUF_TO_STRING.REQ := x > 0;
		BUF_TO_STRING.BUF_FORMAT := TRUE;
		BUF_TO_STRING.BUF_OFFS := DINT#0;
		BUF_TO_STRING.BUF_CNT := DINT#40;
		BUF_TO_STRING.BUFFER := buf;
		BUF_TO_STRING.DST := SHA1_TO_STRH;
		BUF_TO_STRING();
		buf := BUF_TO_STRING.BUFFER;
		SHA1_TO_STRH := BUF_TO_STRING.DST;
	END_FOR;

END_FUNCTION_BLOCK

(* ---- 311-CLEAN.ST ---- *)
FUNCTION_BLOCK CLEAN_Block
	VAR_INPUT
		IN :	STRING;
		CX :	STRING;
	END_VAR

	VAR_OUTPUT
		CLEAN :	STRING;
	END_VAR

	VAR
		pos :	INT;
		stop :	INT;
		char :	STRING;
	END_VAR

	CLEAN := IN;
	stop := LEN(in);
	pos := 1;
	WHILE pos <= stop DO
		char := MID(CLEAN, 1, pos);
		IF FIND(cx,char) > 0 THEN
			pos := pos + 1;
		ELSE
			CLEAN := DELETE(CLEAN, 1, pos);
			stop := stop - 1;
		END_IF;
	END_WHILE;

END_FUNCTION_BLOCK

PROGRAM program0
  VAR
    LocalVar0 : STRING;
    LocalVar1 : STRING;
	LocalOUT  : STRING;
	func_block : CLEAN_Block;
  END_VAR
	func_block.IN  := LocalVar0;
	func_block.CX := LocalVar1;
	func_block();
	LocalOUT := func_block.CLEAN;

END_PROGRAM

CONFIGURATION Config0
  RESOURCE Res0 ON PLC
    TASK task0(INTERVAL := T#20ms,PRIORITY := 0);
    PROGRAM instance0 WITH task0 : program0;
  END_RESOURCE
END_CONFIGURATION

(* ---- 312-COUNT_SUBSTRING.ST ---- *)
FUNCTION_BLOCK COUNT_SUBSTRING_Block
	VAR_INPUT
		SEARCH :	STRING;
		STR :	STRING;
	END_VAR

	VAR_OUTPUT
		COUNT_SUBSTRING :	INT;
	END_VAR

	VAR
		pos :	INT;
		size :	INT;
	END_VAR

	COUNT_SUBSTRING := 0;
	size := LEN(SEARCH);
	REPEAT
	pos := FIND(STR,SEARCH);
	IF pos > 0 THEN
		STR := REPLACE(STR, '', size,pos);
		COUNT_SUBSTRING := COUNT_SUBSTRING + 1;
	END_IF;
	UNTIL pos = 0
	END_REPEAT;
END_FUNCTION_BLOCK

PROGRAM program0
  VAR
	SEARCH :	STRING;
	STR :	STRING;

	COUNT_SUBSTRING :	INT;
	func_block : COUNT_SUBSTRING_Block;
  END_VAR
	func_block.SEARCH  :=SEARCH  ;
	func_block.STR   :=STR   ;

	func_block();
	COUNT_SUBSTRING := func_block.COUNT_SUBSTRING;
END_PROGRAM

CONFIGURATION Config0
  RESOURCE Res0 ON PLC
    TASK task0(INTERVAL := T#20ms,PRIORITY := 0);
    PROGRAM instance0 WITH task0 : program0;
  END_RESOURCE
END_CONFIGURATION

(* ---- 313-CDIV.ST ---- *)
TYPE oscat_complex :
  STRUCT
	re : REAL;
	im : REAL;
  END_STRUCT;
END_TYPE

FUNCTION_BLOCK CDIV_Block

	VAR_INPUT
		X :	oscat_complex;
		Y :	oscat_complex;
	END_VAR

	VAR_OUTPUT
		CDIV :	oscat_complex;
	END_VAR

	VAR
		temp :	REAL;
	END_VAR

	temp := Y.re * Y.re + Y.im * Y.im;
	IF temp = 0.0 THEN CDIV.re := 0.0;CDIV.im := 0.0;RETURN;END_IF;
	CDIV.re := (X.re * Y.re + X.im * Y.im) / temp;
	CDIV.im := (X.im * Y.re - X.re * Y.im) / temp;

END_FUNCTION_BLOCK

PROGRAM program0

	VAR
		X :	oscat_complex;
		Y :	oscat_complex;

		CDIV :	oscat_complex;

		func_block : CDIV_Block;
	END_VAR
	func_block.X := X;
	func_block.Y := Y;
	func_block();
	CDIV := func_block.CDIV;

END_PROGRAM

CONFIGURATION Config0

	RESOURCE Res0 ON PLC
		TASK task0(INTERVAL := T#20ms,PRIORITY := 0);
		PROGRAM instance0 WITH task0 : program0;
	END_RESOURCE

END_CONFIGURATION

(* ---- 314-TO_UML.ST ---- *)
FUNCTION _BYTE_TO_INT:INT
	VAR_INPUT
		IN :	BYTE;
	END_VAR

	_BYTE_TO_INT := USINT_TO_INT(BYTE_TO_USINT(IN));
END_FUNCTION

FUNCTION_BLOCK TO_UML_Block

	VAR_INPUT
		IN :	BYTE;
	END_VAR

	VAR_OUTPUT
		TO_UML :	STRING;
	END_VAR

	CASE _BYTE_TO_INT(in) OF
		196:
			TO_UML := 'Ae';
		214:
			TO_UML := 'Oe';
		220:
			TO_UML := 'Ue';
		223:
			TO_UML := 'ss';
		228:
			TO_UML := 'ae';
		246:
			TO_UML := 'oe';
		252:
			TO_UML := 'ue';
	ELSE
		TO_UML := BYTE_TO_STRING(IN);
	END_CASE;

END_FUNCTION_BLOCK

PROGRAM program0
  VAR
	IN :	BYTE;
	TO_UML :	STRING;
	func_block : TO_UML_Block;
  END_VAR
	func_block.IN  := IN;
	func_block();
	TO_UML := func_block.TO_UML;

END_PROGRAM

CONFIGURATION Config0
	RESOURCE Res0 ON PLC
		TASK task0(INTERVAL := T#20ms,PRIORITY := 0);
		PROGRAM instance0 WITH task0 : program0;
	END_RESOURCE
END_CONFIGURATION

(* ---- 315-ARRAY_MIN.ST ---- *)
TYPE
	oscat_pt_ARRAY: ARRAY [1..100] OF REAL;
END_TYPE

FUNCTION_BLOCK ARRAY_MIN_Block
	VAR_IN_OUT
		PT :	oscat_pt_ARRAY;
	END_VAR

	VAR_INPUT
		SIZE :	UINT;
	END_VAR

	VAR_OUTPUT
		ARRAY_MIN :	REAL;
	END_VAR

	VAR
		i :	INT;
		stop :	INT;
	END_VAR

	stop :=LIMIT_INT(1,UINT_TO_INT(size),1000);

	array_min := pt[1];
	FOR i := 2 TO stop DO
		IF pt[i] < array_min THEN array_min := pt[i]; END_IF;
	END_FOR;

END_FUNCTION_BLOCK
PROGRAM program0
  VAR
    LocalVar0 : oscat_pt_ARRAY;
    LocalVar1 : UINT;
	LocalOUT  : REAL;
	func_block : ARRAY_MIN_Block;
  END_VAR
	func_block.pt := LocalVar0;
	func_block.size := LocalVar1;
	func_block();
	LocalOUT := func_block.ARRAY_MIN;

END_PROGRAM

CONFIGURATION Config0
  RESOURCE Res0 ON PLC
    TASK task0(INTERVAL := T#20ms,PRIORITY := 0);
    PROGRAM instance0 WITH task0 : program0;
  END_RESOURCE
END_CONFIGURATION

(* ---- 316-LOWERCASE.ST ---- *)
FUNCTION_BLOCK LOWERCASE_Block

	VAR_INPUT
		STR :	STRING;
	END_VAR

	VAR_OUTPUT
		LOWERCASE :	STRING;
	END_VAR

	VAR
		char :	BYTE;
		char2 :	BYTE;
		pos :	INT;
		l :	INT;
		str_temp :	STRING;
	END_VAR

	LOWERCASE := str;
	l := LEN(str);
	FOR pos := 1 TO l DO
		char := INT_TO_BYTE(GET_CHAR(str,pos));
		char2 := TO_LOWER(char);
		IF char <> char2 THEN
			str_temp := LOWERCASE;
			LOWERCASE := REPLACE(str_temp,BYTE_TO_STRING(char2,'%c'),1,pos);
		END_IF;
	END_FOR;

END_FUNCTION_BLOCK

PROGRAM program0
  VAR
    OCT : STRING;
    LOWERCASE : STRING;
	func_block : LOWERCASE_Block;
  END_VAR

  	func_block.OCT := '125';
	func_block();
	LOWERCASE := func_block.LOWERCASE;
END_PROGRAM

CONFIGURATION Config0
	RESOURCE Res0 ON PLC
		TASK task0(INTERVAL := T#20ms,PRIORITY := 0);
		PROGRAM instance0 WITH task0 : program0;
	END_RESOURCE
END_CONFIGURATION

(* ---- 318-UPPERCASE.ST ---- *)
FUNCTION_BLOCK UPPERCASE_Block

	VAR_INPUT
		STR :	STRING;
	END_VAR

	VAR_OUTPUT
		UPPERCASE :	STRING;
	END_VAR

	VAR
		char :	BYTE;
		char2 :	BYTE;
		pos :	INT;
		l :	INT;
		str_temp :	STRING;
	END_VAR

	UPPERCASE := str;
	l := LEN(str);
	FOR pos := 1 TO l DO
		char := INT_TO_BYTE(GET_CHAR(str,pos));
		char2 := TO_UPPER(char);
		IF char <> char2 THEN
			str_temp := UPPERCASE;
			UPPERCASE := REPLACE(str_temp,BYTE_TO_STRING(char2,'%c'),1,pos);
		END_IF;
	END_FOR;

END_FUNCTION_BLOCK

PROGRAM program0
	VAR
	    LocalVar1 : STRING;
		LocalOUT  : STRING;
		func_block : UPPERCASE_Block;
  	END_VAR
	func_block.STR := LocalVar1;
	func_block();
	LocalOUT := func_block.UPPERCASE;
END_PROGRAM

CONFIGURATION Config0
  	RESOURCE Res0 ON PLC
    	TASK task0(INTERVAL := T#20ms,PRIORITY := 0);
    	PROGRAM instance0 WITH task0 : program0;
  	END_RESOURCE
END_CONFIGURATION

(* ---- 319-CLICK_CNT.ST ---- *)
FUNCTION_BLOCK CLICK_CNT
	VAR_INPUT
		IN :	BOOL;
		N :	INT;
		TC :	TIME;
	END_VAR

	VAR_OUTPUT
		Q :	BOOL;
	END_VAR

	VAR
		tx :	TP;
		edge :	BOOL;
		cnt :	INT := INT#-1;
	END_VAR

	Q := FALSE;

	IF in AND NOT edge AND NOT tx.q THEN
		cnt := 0;
	ELSIF tx.Q AND NOT IN AND edge THEN
		cnt := cnt + 1;
	ELSIF NOT tx.Q THEN
		Q := cnt=N;
		cnt := -1;
	END_IF;
	edge := IN;
	tx(in := IN, pt := TC);
END_FUNCTION_BLOCK

PROGRAM program0
  VAR
    LocalVar0 : BOOl;
    LocalVar1 : INT;
	LocalVar2 : TIME;
	LocalOUT  : BOOL;
	func_block : CLICK_CNT;
  END_VAR
	func_block.IN  := LocalVar0;
	func_block.N := LocalVar1;
	func_block.TC  := LocalVar2;
	func_block();
	LocalOUT := func_block.Q;

END_PROGRAM

CONFIGURATION Config0
  RESOURCE Res0 ON PLC
    TASK task0(INTERVAL := T#20ms,PRIORITY := 0);
    PROGRAM instance0 WITH task0 : program0;
  END_RESOURCE
END_CONFIGURATION

(* ---- 320-DEL_CHARS.ST ---- *)
FUNCTION_BLOCK DEL_CHARS_Block
	VAR_INPUT
		IN :	STRING;
		CX :	STRING;
	END_VAR

	VAR_OUTPUT
		DEL_CHARS :	STRING;
	END_VAR

	VAR
		pos :	INT;
		stop :	INT;
		char :	STRING;
	END_VAR

	DEL_CHARS := IN;
	stop := LEN(in);
	pos := 1;
	WHILE pos <= stop DO
		char := MID(DEL_CHARS, 1, pos);
		IF FIND(cx,char) > 0 THEN
			DEL_CHARS := DELETE(DEL_CHARS, 1, pos);
			stop := stop - 1;
		ELSE
			pos := pos + 1;
		END_IF;
	END_WHILE;

END_FUNCTION_BLOCK

PROGRAM program0
  VAR
    LocalVar0 : STRING;
	LocalVar1 : STRING;
	LocalOUT  : STRING;
	func_block : DEL_CHARS_Block;
  END_VAR
	func_block.IN := LocalVar0;
	func_block.CX  := LocalVar1;
	func_block();
	LocalOUT := func_block.DEL_CHARS;
END_PROGRAM

CONFIGURATION Config0
  RESOURCE Res0 ON PLC
    TASK task0(INTERVAL := T#20ms,PRIORITY := 0);
    PROGRAM instance0 WITH task0 : program0;
  END_RESOURCE
END_CONFIGURATION

(* ---- 321-FT_MIN_MAX.ST ---- *)
FUNCTION_BLOCK FT_MIN_MAX_Block

  VAR_INPUT
    IN :	REAL;
    RST :	BOOL;
  END_VAR

  VAR_OUTPUT
    MX :	REAL;
    MN :	REAL;
  END_VAR

  VAR
    init :	BOOL;
  END_VAR

  IF (rst = TRUE) OR (init = FALSE) THEN
    mn := in;
    mx := in;
    init := TRUE;
  ELSIF (in < mn) THEN
    mn := in;
  ELSIF (in > mx) THEN
    mx := in;
  END_IF;

END_FUNCTION_BLOCK

PROGRAM program0
  VAR
    IN :	REAL;
    RST :	BOOL;

	  MX :	REAL;
    MN :	REAL;

  	func_block : FT_MIN_MAX_Block;
  END_VAR

	func_block.IN :=IN;
	func_block.RST := RST;
	func_block();
	MX := func_block.MX;
	MN := func_block.MN;

END_PROGRAM

CONFIGURATION Config0

	VAR_GLOBAL
		PLC_TICKS_PER_SEC :	INT;
		PLC_SYS_TICK_CNT :	DINT;
	END_VAR

	RESOURCE Res0 ON PLC
		TASK task0(INTERVAL := T#20ms,PRIORITY := 0);
		PROGRAM instance0 WITH task0 : program0;
	END_RESOURCE

END_CONFIGURATION

(* ---- 322-TRIM1.ST ---- *)
FUNCTION_BLOCK TRIM1

	VAR_INPUT
		STR :	STRING;
	END_VAR

	VAR_OUTPUT
		TRIM3 :	STRING;
	END_VAR

	VAR
		pos :	INT;
		st_temp :	STRING;
	END_VAR

	trim3 := str;
	REPEAT
		pos := FIND(trim3,'  ');
		IF pos > 0 THEN
		st_temp := trim3;
		trim3 := REPLACE(trim3,' ',2,pos);
		END_IF;
	UNTIL pos = 0 END_REPEAT;
	st_temp := LEFT(trim3,1);
	IF EQ_STRING(st_temp,' ') THEN trim3 := DELETE(trim3,1,1); END_IF;
	st_temp := RIGHT(trim3,1);
	IF EQ_STRING(st_temp,' ') THEN trim3 := DELETE(trim3,1,LEN(trim3)); END_IF;

END_FUNCTION_BLOCK

PROGRAM program0
  VAR
	STR :	STRING;

	TRIM3 :	STRING;
	func_block : TRIM1;
  END_VAR
	func_block.STR  :=STR ;
	func_block();
	TRIM3 := func_block.TRIM3;

END_PROGRAM

CONFIGURATION Config0
	RESOURCE Res0 ON PLC
		TASK task0(INTERVAL := T#20ms,PRIORITY := 0);
		PROGRAM instance0 WITH task0 : program0;
	END_RESOURCE
END_CONFIGURATION

(* ---- 323-CATAN.ST ---- *)
TYPE oscat_complex :
  STRUCT
	re : REAL;
	im : REAL;
  END_STRUCT;
END_TYPE

FUNCTION_BLOCK CATAN_Block
	VAR_INPUT
		X :	oscat_complex;
	END_VAR

	VAR_OUTPUT
		CATAN :	oscat_complex;
	END_VAR

	VAR
		r2 :	REAL;
		num :	REAL;
		den :	REAL;
	END_VAR

	r2 := x.re * x.re;
	den := 1.0 - r2 - x.im * x.im;
	CATAN.re := 0.5 * ATAN(2.0 * x.re / den);
	num := x.im + 1.0;
	num := r2 + num * num;
	den := x.im - 1.0;
	den := r2 + den * den;
	CATAN.im := 0.25 * (LN(num)-LN(den));

END_FUNCTION_BLOCK

PROGRAM program0
  VAR
    LocalVar0 : oscat_complex;
	LocalOUT  : oscat_complex;
	func_block : CATAN_Block;
  END_VAR
	func_block.X  := LocalVar0;
	func_block();
	LocalOUT := func_block.CATAN;
END_PROGRAM

CONFIGURATION Config0
  RESOURCE Res0 ON PLC
    TASK task0(INTERVAL := T#20ms,PRIORITY := 0);
    PROGRAM instance0 WITH task0 : program0;
  END_RESOURCE
END_CONFIGURATION

(* ---- 325-_ARRAY_MUL.ST ---- *)
TYPE
	oscat_pt_ARRAY: ARRAY [1..100] OF REAL;
END_TYPE

FUNCTION_BLOCK _ARRAY_MUL2
	VAR_IN_OUT
		PT :	oscat_pt_ARRAY;
	END_VAR
	VAR_INPUT
		SIZE :	UINT;
		X :	REAL;
	END_VAR
	VAR_OUTPUT
		_ARRAY_MUL :	BOOL;
	END_VAR
	VAR
		i :	INT;
		stop :	INT;
	END_VAR

	stop :=LIMIT_INT(1,UINT_TO_INT(size),1000);
	FOR i := 1 TO stop DO
		pt[i] := pt[i] * X;
	END_FOR;
	_ARRAY_MUL := TRUE;

END_FUNCTION_BLOCK

PROGRAM program0
  VAR
    LocalVar0 : oscat_pt_ARRAY;
    LocalVar1 : UINT;
	LocalVar2 : REAL;
	LocalOUT  : BOOL;
	func_block : _ARRAY_MUL2;
  END_VAR
	func_block.pt := LocalVar0;
	func_block.size := LocalVar1;
	func_block.x := LocalVar2;
	func_block();
	LocalOUT := func_block._ARRAY_MUL;

END_PROGRAM

CONFIGURATION Config0
  RESOURCE Res0 ON PLC
    TASK task0(INTERVAL := T#20ms,PRIORITY := 0);
    PROGRAM instance0 WITH task0 : program0;
  END_RESOURCE
END_CONFIGURATION

(* ---- 326-ARRAY_AVG.ST ---- *)
TYPE
	oscat_pt_ARRAY: ARRAY [1..100] OF REAL;
END_TYPE

FUNCTION_BLOCK ARRAY_AVG_Block
	VAR_IN_OUT
		PT :	oscat_pt_ARRAY;
	END_VAR

	VAR_INPUT
		SIZE :	UINT;
	END_VAR

	VAR_OUTPUT
		ARRAY_AVG :	REAL;
	END_VAR

	VAR
		i :	INT;
		stop :	INT;
	END_VAR

	stop :=LIMIT_INT(1,UINT_TO_INT(size),1000);

	array_avg := 0.0;
	FOR i := 1 TO stop DO
		array_avg := array_avg + pt[i];
	END_FOR;
	array_avg := array_avg / INT_TO_REAL(stop);
END_FUNCTION_BLOCK

PROGRAM program0
  VAR
    LocalVar0 : oscat_pt_ARRAY;
    LocalVar1 : UINT;
	LocalOUT  : REAL;
	func_block : ARRAY_AVG_Block;
  END_VAR
	func_block.pt := LocalVar0;
	func_block.size := LocalVar1;
	func_block();
	LocalOUT := func_block.ARRAY_AVG;

END_PROGRAM

CONFIGURATION Config0
  RESOURCE Res0 ON PLC
    TASK task0(INTERVAL := T#20ms,PRIORITY := 0);
    PROGRAM instance0 WITH task0 : program0;
  END_RESOURCE
END_CONFIGURATION

(* ---- 327-CATANH.ST ---- *)
TYPE oscat_complex :
  STRUCT
	re : REAL;
	im : REAL;
  END_STRUCT;
END_TYPE

FUNCTION_BLOCK CATANH_Block
	VAR_INPUT
		X :	oscat_complex;
	END_VAR

	VAR_OUTPUT
		CATANH :	oscat_complex;
	END_VAR

	VAR
		i2 :	REAL;
		num :	REAL;
		den :	REAL;
	END_VAR

	i2 := x.im * x.im;
	num := 1.0 + x.re;
	num := i2 + num * num;
	den := 1.0 - x.re;
	den := i2 + den * den;
	CATANH.re := 0.25 * (LN(num) - LN(den));
	den := 1.0 - x.re * x.re - i2;
	CATANH.im := 0.5 * ATAN(2.0 * x.im / den);

END_FUNCTION_BLOCK

PROGRAM program0
  VAR
    LocalVar0 : oscat_complex;
	LocalOUT  : oscat_complex;
	func_block : CATANH_Block;
  END_VAR
	func_block.X  := LocalVar0;
	func_block();
	LocalOUT := func_block.CATANH;
END_PROGRAM

CONFIGURATION Config0
  RESOURCE Res0 ON PLC
    TASK task0(INTERVAL := T#20ms,PRIORITY := 0);
    PROGRAM instance0 WITH task0 : program0;
  END_RESOURCE
END_CONFIGURATION

(* ---- 328-IRTRANS_RCV_1.ST ---- *)
FUNCTION_BLOCK IRTRANS_RCV_1_Block

	VAR_INPUT
		CMD :	BOOL;
		DEV_CODE :	STRING;
		KEY_CODE :	STRING;
	END_VAR

	VAR_OUTPUT
		Q :	BOOL;
	END_VAR

	VAR_IN_OUT
		DEV :	STRING;
		KEY :	STRING;
	END_VAR

	Q := cmd AND EQ_STRING(dev_code,dev) AND EQ_STRING(key_code,key);

END_FUNCTION_BLOCK

PROGRAM program0
	VAR
		CMD :	BOOL;
		DEV :	STRING;
		KEY :	STRING;
		DEV_CODE :	STRING;
		KEY_CODE :	STRING;
		Q :	BOOL;

		func_block : IRTRANS_RCV_1_Block;
	END_VAR
	func_block.CMD := CMD;
	func_block.DEV := DEV;
	func_block.KEY := KEY;
	func_block.DEV_CODE := DEV_CODE;
	func_block.KEY_CODE := KEY_CODE;

	func_block();
	DEV  := func_block.DEV;
	KEY  := func_block.KEY;
	Q  := func_block.Q;

END_PROGRAM

CONFIGURATION Config0

  	RESOURCE Res0 ON PLC
    	TASK task0(INTERVAL := T#20ms,PRIORITY := 0);
    	PROGRAM instance0 WITH task0 : program0;
  	END_RESOURCE

END_CONFIGURATION

(* ---- 329-BUFFER_CLEAR.ST ---- *)
TYPE
	oscat_arb_0_249 			  : ARRAY [0..249] 	OF BYTE;
END_TYPE

FUNCTION_BLOCK _BUFFER_CLEAR
	VAR_IN_OUT
		PT :	oscat_arb_0_249;
	END_VAR

	VAR_INPUT
		SIZE :	UINT;
	END_VAR

	VAR_OUTPUT
		BUFFER_CLEAR :	BOOL;
	END_VAR

	VAR
		err :	INT;
		result :	WORD;
	END_VAR

	result := MEMSET(err,BYTE#00,UINT_TO_DINT(size),pt[0]);
	BUFFER_CLEAR := (err = 0);

END_FUNCTION_BLOCK

PROGRAM program0
	VAR
	    LocalVar1 : oscat_arb_0_249;
		LocalVar2 : UINT;
		LocalOUT  : BOOL;
		func_block : _BUFFER_CLEAR;
  	END_VAR
	func_block.PT := LocalVar1;
	func_block.SIZE := LocalVar2;
	func_block();
	LocalOUT := func_block.BUFFER_CLEAR;
END_PROGRAM

CONFIGURATION Config0
	VAR_GLOBAL
		PLC_TICKS_PER_SEC :	INT;
		PLC_SYS_TICK_CNT :	DINT;
	END_VAR

  	RESOURCE Res0 ON PLC
    	TASK task0(INTERVAL := T#20ms,PRIORITY := 0);
    	PROGRAM instance0 WITH task0 : program0;
  	END_RESOURCE
END_CONFIGURATION

(* ---- 330-OCT_TO_BYTE.ST ---- *)
FUNCTION_BLOCK OCT_TO_BYTE_Block
	VAR_INPUT
		OCT :	STRING;
	END_VAR

	VAR_OUTPUT
		OCT_TO_BYTE :	BYTE;
	END_VAR

	VAR
		i :	INT;
		stop :	INT;
		X :	INT;
	END_VAR

	OCT_TO_BYTE := BYTE#0;
	stop := LEN(oct);
	FOR I := 1 TO stop DO
		(* read the first character and subtract 48 to get value in decimal 0 = 48 *)
		X := GET_CHAR(oct,I);
		(* calculate the value of the digit *)
		IF X > 47 AND x < 56 THEN
			OCT_TO_BYTE := SHL_BYTE(OCT_TO_BYTE,3) OR INT_TO_BYTE(X - 48);
		END_IF;
	END_FOR;

END_FUNCTION_BLOCK

PROGRAM program0
  VAR
    OCT : STRING;
    OCT_TO_BYTE : BYTE;
	func_block : OCT_TO_BYTE_Block;
  END_VAR

  	func_block.OCT := '125';
	func_block();
	OCT_TO_BYTE := func_block.OCT_TO_BYTE;
END_PROGRAM

CONFIGURATION Config0
	RESOURCE Res0 ON PLC
		TASK task0(INTERVAL := T#20ms,PRIORITY := 0);
		PROGRAM instance0 WITH task0 : program0;
	END_RESOURCE
END_CONFIGURATION

(* ---- 332-HYST_3.ST ---- *)
FUNCTION_BLOCK HYST_3_Block

	VAR_INPUT
		IN :	REAL;
		HYST :	REAL;
		VAL1 :	REAL;
		VAL2 :	REAL;
	END_VAR

	VAR_OUTPUT
		Q1 :	BOOL;
		Q2 :	BOOL;
	END_VAR

	VAR
		X :	REAL;
	END_VAR

	X := hyst * 0.5;
	IF in < val1 - X THEN
		q1 := TRUE;
	ELSIF in > val1 + X THEN
		q1 := FALSE;
	END_IF;
	IF in < val2 - X THEN
		q2 := FALSE;
	ELSIF in > val2 + X THEN
		q2 := TRUE;
	END_IF;

END_FUNCTION_BLOCK

PROGRAM program0
	VAR
		IN :	REAL;
		HYST :	REAL;
		VAL1 :	REAL;
		VAL2 :	REAL;
		Q1 :	BOOL;
		Q2 :	BOOL;
		func_block : HYST_3_Block;
	END_VAR
	func_block.IN := IN;
	func_block.HYST := HYST;
	func_block.VAL1 := VAL1;
	func_block.VAL2 := VAL2;
	func_block();
	Q1  := func_block.Q1;
	Q2  := func_block.Q2;
END_PROGRAM

CONFIGURATION Config0
	RESOURCE Res0 ON PLC
		TASK task0(INTERVAL := T#20ms,PRIORITY := 0);
		PROGRAM instance0 WITH task0 : program0;
	END_RESOURCE
END_CONFIGURATION

(* ---- 333-_ARRAY_INIT.ST ---- *)
TYPE
	oscat_pt_ARRAY: ARRAY [1..100] OF REAL;
END_TYPE

FUNCTION_BLOCK _ARRAY_INIT2

	VAR_IN_OUT
		PT :	oscat_pt_ARRAY;
	END_VAR

	VAR_INPUT
		SIZE :	UINT;
		INIT :	REAL;
	END_VAR

	VAR_OUTPUT
		_ARRAY_INIT:	BOOL;
	END_VAR

	VAR
		i :	INT;
		stop :	INT;
	END_VAR

	stop :=LIMIT_INT(1,UINT_TO_INT(size),1000);

	FOR i := 1 TO stop DO
		pt[i] := init;
	END_FOR;
	_ARRAY_INIT := TRUE;

END_FUNCTION_BLOCK

PROGRAM program0
  VAR
    LocalVar0 : oscat_pt_ARRAY;
    LocalVar1 : UINT;
	LocalVar2 : REAL;
	LocalOUT  : BOOL;
	func_block: _ARRAY_INIT2;
  END_VAR
  func_block.pt := LocalVar0;
  func_block.size := LocalVar1;
  func_block.init := LocalVar2;
  func_block();
  LocalOUT := func_block._ARRAY_INIT;
END_PROGRAM

CONFIGURATION Config0
  RESOURCE Res0 ON PLC
    TASK task0(INTERVAL := T#20ms,PRIORITY := 0);
    PROGRAM instance0 WITH task0 : program0;
  END_RESOURCE
END_CONFIGURATION

(* ---- 337-HYST.ST ---- *)
FUNCTION_BLOCK HYST_Block

	VAR_INPUT
		IN :	REAL;
		_ON :	REAL;
		OFF :	REAL;
	END_VAR

	VAR_OUTPUT
		Q :	BOOL;
		WIN :	BOOL;
	END_VAR

	IF _ON >= OFF THEN
		IF IN < OFF THEN
			Q := FALSE;
			WIN := FALSE;
		ELSIF  IN > _ON THEN
			Q := TRUE;
			WIN := FALSE;
		ELSE
			WIN := TRUE;
		END_IF;
	ELSE
		IF IN > OFF THEN
			Q := FALSE;
			WIN := FALSE;
		ELSIF  IN < _ON THEN
			Q := TRUE;
			WIN := FALSE;
		ELSE
			WIN := TRUE;
		END_IF;
	END_IF;

END_FUNCTION_BLOCK

PROGRAM program0
	VAR
		IN :	REAL;
		_ON :	REAL;
		OFF :	REAL;
		Q :	BOOL;
		WIN :	BOOL;
		func_block : HYST_Block;
	END_VAR
	func_block.IN := IN;
	func_block._ON := _ON;
	func_block.OFF := OFF ;
	func_block();
	Q  := func_block.Q;
	WIN  := func_block.WIN;
END_PROGRAM

CONFIGURATION Config0
	RESOURCE Res0 ON PLC
		TASK task0(INTERVAL := T#20ms,PRIORITY := 0);
		PROGRAM instance0 WITH task0 : program0;
	END_RESOURCE
END_CONFIGURATION

(* ---- 338-SETUP_CHARNAMES.ST ---- *)
TYPE
  oscat_CHARNAMES	: ARRAY [1..11] OF STRING;
END_TYPE

FUNCTION_BLOCK SETUP_CHARNAMES_Block

	VAR_IN_OUT
		CHARNAMES :	oscat_CHARNAMES;
	END_VAR

	VAR
		init :	BOOL;
	END_VAR

	IF init THEN RETURN; END_IF;

	init := TRUE;

	CHARNAMES[01] := '123';
	CHARNAMES[02] := '456';
	CHARNAMES[03] := 'zgsdafasf';
	CHARNAMES[04] := 'sadfsdfa';
	CHARNAMES[05] := 'asdfdsafdfds';
	CHARNAMES[06] := 'sadfsdfsdf';
	CHARNAMES[07] := 'sfsfdfdddd';
	CHARNAMES[08] := 'dddddted';
	CHARNAMES[10] := 'wer';
	CHARNAMES[11] := 'werwer';

END_FUNCTION_BLOCK

PROGRAM program0

	VAR
		CHARNAMES :	oscat_CHARNAMES;
		func_block : SETUP_CHARNAMES_Block;
  	END_VAR
	func_block.CHARNAMES  :=CHARNAMES;
	func_block();
	CHARNAMES := func_block.CHARNAMES;

END_PROGRAM

CONFIGURATION Config0

	RESOURCE Res0 ON PLC
		TASK task0(INTERVAL := T#20ms,PRIORITY := 0);
		PROGRAM instance0 WITH task0 : program0;
	END_RESOURCE

END_CONFIGURATION

(* ---- 339-IS_SORTED.ST ---- *)
TYPE
	oscat_pt_ARRAY: ARRAY [1..100] OF REAL;
END_TYPE

FUNCTION_BLOCK IS_SORTED_Block

	VAR_IN_OUT
		PT :	oscat_pt_ARRAY;
	END_VAR

	VAR_INPUT
		SIZE :	UINT;
	END_VAR

	VAR_OUTPUT
		IS_SORTED :	BOOL;
	END_VAR

	VAR
		i :	INT;
		i2 :	INT;
		stop :	INT;
	END_VAR

	stop :=LIMIT_INT(1,UINT_TO_INT(size),1000);
	stop := stop -1;
	FOR i := 1 TO stop DO
		i2 := i+1;
		IF pt[i] > pt[i2] THEN
			IS_SORTED := FALSE;
			RETURN;
		END_IF;
	END_FOR;

	IS_SORTED := TRUE;

END_FUNCTION_BLOCK

PROGRAM program0

	VAR
		SIZE :	UINT;
		PT :	oscat_pt_ARRAY;
		IS_SORTED :	BOOL;
		func_block : IS_SORTED_Block;
	END_VAR
	func_block.SIZE := SIZE;
	func_block.PT := PT;
	func_block();
	PT := func_block.PT;
	IS_SORTED := func_block.IS_SORTED;

END_PROGRAM

CONFIGURATION Config0

	RESOURCE Res0 ON PLC
		TASK task0(INTERVAL := T#20ms,PRIORITY := 0);
		PROGRAM instance0 WITH task0 : program0;
	END_RESOURCE

END_CONFIGURATION

(* ---- 340-REAL_TO_DW.ST ---- *)
FUNCTION_BLOCK REAL_TO_DW_Block
  VAR_INPUT
    X :	REAL;
  END_VAR

  VAR_OUTPUT
    REAL_TO_DW :	DWORD;
  END_VAR

  VAR
    REAL_TO_BUF :	REAL_TO_BUF;
    i :	INT;
  END_VAR

  FOR I := 0 TO 1 DO
    REAL_TO_BUF.REQ        := I > 0;
    REAL_TO_BUF.BUF_FORMAT := FALSE;
    REAL_TO_BUF.BUF_OFFS   := DINT#0;
    REAL_TO_BUF.BUF_CNT    := DINT#4;
    REAL_TO_BUF.SRC        := X;
    REAL_TO_BUF.BUFFER     := REAL_TO_DW;
    REAL_TO_BUF();
    X          := REAL_TO_BUF.SRC;
    REAL_TO_DW := REAL_TO_BUF.BUFFER;
  END_FOR;
END_FUNCTION_BLOCK

PROGRAM program0
  VAR
    LocalVar0 : REAL;
    LocalOUT  : DWORD;
    func_block : REAL_TO_DW_Block;
  END_VAR
	func_block.X  := LocalVar0;
	func_block();
	LocalOUT := func_block.REAL_TO_DW;

END_PROGRAM

CONFIGURATION Config0
  RESOURCE Res0 ON PLC
    TASK task0(INTERVAL := T#20ms,PRIORITY := 0);
    PROGRAM instance0 WITH task0 : program0;
  END_RESOURCE
END_CONFIGURATION

(* ---- 342-BIN_TO_BYTE.ST ---- *)
TYPE
  oscat_STRING12              : STRING(12);
END_TYPE

FUNCTION_BLOCK BIN_TO_BYTE_Block
	VAR_INPUT
		BIN :	oscat_STRING12;
	END_VAR

	VAR_OUTPUT
		BIN_TO_BYTE :	BYTE;
	END_VAR

	VAR
		i :	INT;
		stop :	INT;
		X :	INT;
	END_VAR

	BIN_TO_BYTE := BYTE#0;
	stop := LEN(bin);
	FOR I := 1 TO LEN(BIN) DO
		X := GET_CHAR(BIN,I);
		(* calculate the value of the digit *)
		IF X = 48 THEN
			BIN_TO_BYTE := SHL_BYTE(BIN_TO_BYTE,1);
		ELSIF X = 49 THEN
			BIN_TO_BYTE := SHL_BYTE(BIN_TO_BYTE,1) OR BYTE#1;
		END_IF;
	END_FOR;

END_FUNCTION_BLOCK

PROGRAM program0
  VAR
    LocalVar0 : oscat_STRING12;
	LocalOUT  : BYTE;
	func_block : BIN_TO_BYTE_Block;
  END_VAR
	func_block.BIN := LocalVar0;
	func_block();
	LocalOUT := func_block.BIN_TO_BYTE;

END_PROGRAM

CONFIGURATION Config0
  RESOURCE Res0 ON PLC
    TASK task0(INTERVAL := T#20ms,PRIORITY := 0);
    PROGRAM instance0 WITH task0 : program0;
  END_RESOURCE
END_CONFIGURATION

(* ---- 343-CALIBRATE.ST ---- *)
FUNCTION_BLOCK CALIBRATE
	VAR_INPUT
		X :	REAL;
		CO :	BOOL;
		CS :	BOOL;
		Y_OFFSET :	REAL;
		Y_SCALE :	REAL;
	END_VAR

	VAR_OUTPUT
		Y :	REAL;
	END_VAR

	VAR RETAIN
		offset :	REAL;
		Scale :	REAL := 1.0;
	END_VAR

	IF CO THEN
		OFFSET := Y_Offset - X;
	ELSIF CS THEN
		SCALE := Y_scale / (X + OFFSET);
	END_IF;
	Y := (X + OFFSET) * SCALE;

END_FUNCTION_BLOCK

PROGRAM program0
  VAR
    LocalVar0 : REAL;
    LocalVar1 : BOOL;
	LocalVar2 : BOOL;
	LocalVar3 : REAL;
	LocalVar4 : REAL;
	LocalOUT  : REAL;
	func_block : CALIBRATE;
  END_VAR
	func_block.X  := LocalVar0;
	func_block.CO := LocalVar1;
	func_block.CS  := LocalVar2;
	func_block.Y_OFFSET := LocalVar3;
	func_block.Y_SCALE := LocalVar4;
	func_block();
	LocalOUT := func_block.Y;

END_PROGRAM

CONFIGURATION Config0
  RESOURCE Res0 ON PLC
    TASK task0(INTERVAL := T#20ms,PRIORITY := 0);
    PROGRAM instance0 WITH task0 : program0;
  END_RESOURCE
END_CONFIGURATION

(* ---- 344-FINDP.ST ---- *)
FUNCTION_BLOCK FINDP_Block

	VAR_INPUT
		STR :	STRING;
		SRC :	STRING;
		POS :	INT;
	END_VAR

	VAR_OUTPUT
		FINDP :	INT;
	END_VAR

	VAR
		i :	INT;
		ls :	INT;
		lx :	INT;
		stp :	INT;
		st_tmp :	STRING;
	END_VAR

	ls := LEN(str);
	lx := LEN(src);
	IF ls < lx OR lx = 0 THEN RETURN; END_IF;
	stp := ls - lx + 1;
	FOR i := MAX(pos,1) TO stp DO
		st_tmp := MID(str,lx,i);
		IF EQ_STRING(st_tmp,src) THEN
			FINDP := i;
			RETURN;
		END_IF;
	END_FOR;
	FINDP := 0;

END_FUNCTION_BLOCK

PROGRAM program0

	VAR
		STR :	STRING;
		SRC :	STRING;
		POS :	INT;

        FINDP :	INT;
		func_block : FINDP_Block;
	END_VAR
		func_block.STR := STR;
		func_block.SRC := SRC;
		func_block.POS := POS;
		func_block();
		FINDP := func_block.FINDP;

END_PROGRAM

CONFIGURATION Config0

	RESOURCE Res0 ON PLC
		TASK task0(INTERVAL := T#20ms,PRIORITY := 0);
		PROGRAM instance0 WITH task0 : program0;
	END_RESOURCE

END_CONFIGURATION

(* ---- 345-SETUP_LOCATION.ST ---- *)
TYPE
	oscat_LOCATION_ELEMENTS	: ARRAY [1..5] OF INT;
END_TYPE

TYPE oscat_LOCATION:
  STRUCT
    DEFAULT 	: INT;
	LMAX    	: INT;
	LANGUAGE	: oscat_LOCATION_ELEMENTS;
  END_STRUCT;
END_TYPE

FUNCTION_BLOCK SETUP_LOCATION_Block
	VAR_IN_OUT
		LOCATION :	oscat_LOCATION;
	END_VAR

	VAR
		init :	BOOL;
	END_VAR

	IF init THEN RETURN; END_IF;
	init := TRUE;

	LOCATION.DEFAULT  := 1;
	LOCATION.LMAX := 5;

	LOCATION.LANGUAGE[1] := 2;
	LOCATION.LANGUAGE[2] := 2;
	LOCATION.LANGUAGE[3] := 3;
	LOCATION.LANGUAGE[4] := 2;
	LOCATION.LANGUAGE[5] := 2;

END_FUNCTION_BLOCK

PROGRAM program0
	VAR
		LOCATION :	oscat_LOCATION;
		func_block : SETUP_LOCATION_Block;
  	END_VAR
	func_block.LOCATION  :=LOCATION;
	func_block();
	LOCATION := func_block.LOCATION;
END_PROGRAM

CONFIGURATION Config0
	RESOURCE Res0 ON PLC
		TASK task0(INTERVAL := T#20ms,PRIORITY := 0);
		PROGRAM instance0 WITH task0 : program0;
	END_RESOURCE
END_CONFIGURATION

(* ---- 346-SPEED.ST ---- *)
FUNCTION_BLOCK SPEED_Block

	VAR_INPUT
		MS :	REAL;
		KMH :	REAL;
		KN :	REAL;
		MH :	REAL;
	END_VAR

	VAR_OUTPUT
		YMS :	REAL;
		YKMH :	REAL;
		YKN :	REAL;
		YMH :	REAL;
	END_VAR

	Yms := ms +
			kmh * 0.27777777777778 +
			kn * 0.5144444 +
			mh * 0.44704;
	Ykmh := Yms * 3.6;
	Ykn := Yms * 1.94384466037535;
	Ymh := Yms * 2.23693629205440;

END_FUNCTION_BLOCK

PROGRAM program0

	VAR
		MS :	REAL;
		KMH :	REAL;
		KN :	REAL;
		MH :	REAL;
		YMS :	REAL;
		YKMH :	REAL;
		YKN :	REAL;
		YMH :	REAL;
		func_block : SPEED_Block;
	END_VAR
		func_block.MS  :=MS;
		func_block.KMH  :=KMH;
		func_block.KN  :=KN;
		func_block.MH  :=MH;
		func_block();
		YMS := func_block.YMS;
		YKMH := func_block.YKMH;
		YKN := func_block.YKN;
		YMH := func_block.YMH;

	END_PROGRAM

CONFIGURATION Config0

	RESOURCE Res0 ON PLC
		TASK task0(INTERVAL := T#20ms,PRIORITY := 0);
		PROGRAM instance0 WITH task0 : program0;
	END_RESOURCE

END_CONFIGURATION

(* ---- 347-TREND_DW.ST ---- *)
FUNCTION_BLOCK TREND_DW
	VAR_INPUT
		X :	DWORD;
	END_VAR
	VAR_OUTPUT
		Q :	BOOL;
		TU :	BOOL;
		TD :	BOOL;
		D :	DWORD;
	END_VAR

	VAR
		LAST_X :	DWORD;
	END_VAR

	IF X > last_X THEN
		TU := TRUE;
		TD := FALSE;
		D := UDINT_TO_DWORD(DWORD_TO_UDINT(X) - DWORD_TO_UDINT(last_X));
		Q := TRUE;
	ELSIF X < last_X THEN
		TD := TRUE;
		TU := FALSE;
		D := UDINT_TO_DWORD(DWORD_TO_UDINT(last_X) - DWORD_TO_UDINT(X));
		Q := FALSE;
	ELSE
		TU := FALSE;
		TD := FALSE;
		D := DWORD#0;
	END_IF;
	last_X := X;
END_FUNCTION_BLOCK

PROGRAM program0
  VAR
	X :	DWORD;
	Q :	BOOL;
	TU :	BOOL;
	TD :	BOOL;
	D :	DWORD;
	func_block : TREND_DW;
  END_VAR
	func_block.X  :=X ;
	func_block();
	Q := func_block.Q;
	TU := func_block.TU;
	TD := func_block.TD;
	D := func_block.D;
END_PROGRAM

CONFIGURATION Config0
	RESOURCE Res0 ON PLC
		TASK task0(INTERVAL := T#20ms,PRIORITY := 0);
		PROGRAM instance0 WITH task0 : program0;
	END_RESOURCE
END_CONFIGURATION

(* ---- 348-V3_ZANG.ST ---- *)
TYPE oscat_vector_3:
  STRUCT
	X : REAL;
	Y : REAL;
	Z : REAL;
  END_STRUCT;
END_TYPE

FUNCTION_BLOCK V3_ABS_Block

	VAR_INPUT
		A :	oscat_vector_3;
	END_VAR

	VAR_OUTPUT
		V3_ABS :	REAL;
	END_VAR

	V3_ABS := SQRT(A.X * A.X + A.Y * A.Y + A.Z * A.Z);

END_FUNCTION_BLOCK

FUNCTION_BLOCK V3_ZANG_Block
	VAR_INPUT
		A :	oscat_vector_3;
	END_VAR

	VAR_OUTPUT
		V3_ZANG :	REAL;
	END_VAR

	VAR
		la :	REAL;
		V3_ABS :	V3_ABS_Block;
	END_VAR

	V3_ABS(A:=A);
	la:=V3_ABS.V3_ABS;

	IF la > 0.0 THEN
		V3_ZANG := ACOS(A.Z / la);
	ELSE
		V3_ZANG := 0.0;
	END_IF;

END_FUNCTION_BLOCK

PROGRAM program0
  	VAR
		A :	oscat_vector_3;
		V3_ZANG :	REAL;
		func_block : V3_ZANG_Block;
  	END_VAR
	func_block.A := A;
	func_block();
	V3_ZANG := func_block.V3_ZANG;
END_PROGRAM

CONFIGURATION Config0
  RESOURCE Res0 ON PLC
    TASK task0(INTERVAL := T#20ms,PRIORITY := 0);
    PROGRAM instance0 WITH task0 : program0;
  END_RESOURCE
END_CONFIGURATION

(* ---- 349-V3_YANG.ST ---- *)
TYPE oscat_vector_3:
  	STRUCT
		X : REAL;
		Y : REAL;
		Z : REAL;
  	END_STRUCT;
END_TYPE

FUNCTION_BLOCK V3_ABS_Block

	VAR_INPUT
		A :	oscat_vector_3;
	END_VAR

	VAR_OUTPUT
		V3_ABS :	REAL;
	END_VAR

	V3_ABS := SQRT(A.X * A.X + A.Y * A.Y + A.Z * A.Z);

END_FUNCTION_BLOCK

FUNCTION_BLOCK V3_YANG_Block
	VAR_INPUT
		A :	oscat_vector_3;
	END_VAR

	VAR_OUTPUT
		V3_YANG :	REAL;
	END_VAR

	VAR
		la :	REAL;
		V3_ABS :	V3_ABS_Block;
	END_VAR

	V3_ABS(A:=A);
	la:=V3_ABS.V3_ABS;

	IF la > 0.0 THEN
		V3_YANG := ACOS(A.Y / la);
	ELSE
		V3_YANG := 0.0;
	END_IF;

END_FUNCTION_BLOCK

PROGRAM program0
  	VAR
		A :	oscat_vector_3;
		V3_YANG :	REAL;
		func_block : V3_YANG_Block;
  	END_VAR
	func_block.A := A;
	func_block();
	V3_YANG := func_block.V3_YANG;
END_PROGRAM

CONFIGURATION Config0
  RESOURCE Res0 ON PLC
    TASK task0(INTERVAL := T#20ms,PRIORITY := 0);
    PROGRAM instance0 WITH task0 : program0;
  END_RESOURCE
END_CONFIGURATION

(* ---- 350-_INSERT80.ST ---- *)
FUNCTION_BLOCK _INSERT80

    VAR_INPUT
        IN1 :	STRING;
        IN2 :	STRING;
        P :	INT;
    END_VAR

    VAR_OUTPUT
        _INSERT :	STRING;
    END_VAR

    VAR
        size :	INT;
    END_VAR

    size := LEN(IN1);
    IF size + LEN(IN2) <= 80 THEN
        P := LIMIT(0,P,size);
        IF P = 0 THEN
            _INSERT := CONCAT(IN2,IN1);
        ELSE
            _INSERT := INSERT(IN1, IN2, P);
        END_IF;
    END_IF;

END_FUNCTION_BLOCK

PROGRAM program0
	VAR
	    LocalVar1 : STRING;
        LocalVar2 : STRING;
        LocalVar3 : INT;
		LocalOUT  : STRING;
		func_block : _INSERT80;
  	END_VAR
	func_block.IN1 := LocalVar1;
    func_block.IN2 := LocalVar2;
    func_block.P := LocalVar3;
	func_block();
	LocalOUT := func_block._INSERT;
END_PROGRAM

CONFIGURATION Config0
  	RESOURCE Res0 ON PLC
    	TASK task0(INTERVAL := T#20ms,PRIORITY := 0);
    	PROGRAM instance0 WITH task0 : program0;
  	END_RESOURCE
END_CONFIGURATION

(* ---- 351-PERIOD2.ST ---- *)
TYPE
	oscat_PERIOD2_Y             : ARRAY [0..1]    OF UDINT;
	oscat_PERIOD2_X             : ARRAY [0..3]    OF oscat_PERIOD2_Y := [0, 0, 0, 0];
END_TYPE

FUNCTION_BLOCK PERIOD2_Block

	VAR_INPUT
		DP :	oscat_PERIOD2_X;
		DX :	UDINT;
	END_VAR

	VAR_OUTPUT
		PERIOD2 :	BOOL;
	END_VAR

	(*@KEY@: WORKSHEET
	NAME: PERIOD2
	IEC_LANGUAGE: ST
	*)
	PERIOD2 := 	(DX >= DP[0][0] AND DX <= DP[0][1]) OR
				(DX >= DP[1][0] AND DX <= DP[1][1]) OR
				(DX >= DP[2][0] AND DX <= DP[2][1]) OR
				(DX >= DP[3][0] AND DX <= DP[3][1]);

END_FUNCTION_BLOCK

PROGRAM program0

	VAR
		DP :	oscat_PERIOD2_X;
		DX :	UDINT;

		PERIOD2 :	BOOL;
		func_block : PERIOD2_Block;
  	END_VAR

	func_block.DP := DP;
	func_block.DX := DX;
	func_block();
	PERIOD2 := func_block.PERIOD2;

END_PROGRAM

CONFIGURATION Config0

  	RESOURCE Res0 ON PLC
    	TASK task0(INTERVAL := T#20ms,PRIORITY := 0);
    	PROGRAM instance0 WITH task0 : program0;
  	END_RESOURCE

END_CONFIGURATION

(* ---- 352-V3_XANG.ST ---- *)
TYPE oscat_vector_3 :
	STRUCT
		X : REAL;
		Y : REAL;
		Z : REAL;
	END_STRUCT;
END_TYPE

FUNCTION_BLOCK V3_ABS_Block

	VAR_INPUT
		A :	oscat_vector_3;
	END_VAR

	VAR_OUTPUT
		V3_ABS :	REAL;
	END_VAR

	V3_ABS := SQRT(A.X * A.X + A.Y * A.Y + A.Z * A.Z);

END_FUNCTION_BLOCK

FUNCTION_BLOCK V3_XANG_Block

	VAR_INPUT
		A :	oscat_vector_3;
	END_VAR

	VAR_OUTPUT
		V3_XANG :	REAL;
	END_VAR

	VAR
		la :	REAL;
		V3_ABS :	V3_ABS_Block;
	END_VAR

	V3_ABS(A:=A);
	la:=V3_ABS.V3_ABS;

	IF la > 0.0 THEN
		V3_XANG := ACOS(A.X / la);
	ELSE
		V3_XANG := 0.0;
	END_IF;

END_FUNCTION_BLOCK

PROGRAM program0
  	VAR
		A :	oscat_vector_3;
		V3_XANG :	REAL;
		func_block : V3_XANG_Block;
  	END_VAR
	func_block.A := A;
	func_block();
	V3_XANG := func_block.V3_XANG;
END_PROGRAM

CONFIGURATION Config0
  RESOURCE Res0 ON PLC
    TASK task0(INTERVAL := T#20ms,PRIORITY := 0);
    PROGRAM instance0 WITH task0 : program0;
  END_RESOURCE
END_CONFIGURATION

(* ---- 353-ARRAY_HAV.ST ---- *)
TYPE
	oscat_pt_ARRAY: ARRAY [1..100] OF REAL;
END_TYPE

FUNCTION_BLOCK ARRAY_HAV_Block
	VAR_IN_OUT
		PT :	oscat_pt_ARRAY;
	END_VAR

	VAR_INPUT
		SIZE :	UINT;
	END_VAR

	VAR_OUTPUT
		ARRAY_HAV :	REAL;
	END_VAR

	VAR
		i :	INT;
		stop :	INT;
	END_VAR

	stop :=LIMIT_INT(1,UINT_TO_INT(size),1000);
	ARRAY_HAV := 0.0;
	FOR i := 1 TO stop DO
		IF pt[i] <> 0.0 THEN
			ARRAY_HAV := ARRAY_HAV + 1.0/pt[i];
		ELSE
			ARRAY_HAV := 0.0;
			RETURN;
		END_IF;
	END_FOR;
	ARRAY_HAV := INT_TO_REAL(stop) / ARRAY_HAV;
END_FUNCTION_BLOCK

PROGRAM program0
  VAR
    LocalVar0 : oscat_pt_ARRAY;
    LocalVar1 : UINT;
	LocalOUT  : REAL;
	func_block : ARRAY_HAV_Block;
  END_VAR
	func_block.pt := LocalVar0;
	func_block.size := LocalVar1;
	func_block();
	LocalOUT := func_block.ARRAY_HAV;

END_PROGRAM

CONFIGURATION Config0
  RESOURCE Res0 ON PLC
    TASK task0(INTERVAL := T#20ms,PRIORITY := 0);
    PROGRAM instance0 WITH task0 : program0;
  END_RESOURCE
END_CONFIGURATION

(* ---- 354-CSIN.ST ---- *)
TYPE oscat_complex :
  STRUCT
	re : REAL;
	im : REAL;
  END_STRUCT;
END_TYPE

FUNCTION COSH:REAL
	VAR_INPUT
		X :	REAL;
	END_VAR

	VAR
		t :	REAL;
	END_VAR

	T := EXP(X);
	COSH := (1.0 / T + T) * 0.5;
END_FUNCTION

FUNCTION SINH:REAL
	VAR_INPUT
		X :	REAL;
	END_VAR

	IF ABS(x) < 2.0E-3 THEN
		SINH := X;
	ELSE
		SINH := (EXP(x) - EXP(-x)) * 0.5;
	END_IF;
END_FUNCTION

FUNCTION_BLOCK CSIN_Block
	VAR_INPUT
		X :	oscat_complex;
	END_VAR

	VAR_OUTPUT
		CSIN :	oscat_complex;
	END_VAR

	CSIN.re := cosH(X.im) * SIN(X.re);
	CSIN.im := sinH(X.im) * COS(X.re);
END_FUNCTION_BLOCK

PROGRAM program0
  VAR
    LocalVar0 : oscat_complex;
	LocalOUT  : oscat_complex;
	func_block : CSIN_Block;
  END_VAR
	func_block.X  := LocalVar0;
	func_block();
	LocalOUT := func_block.CSIN;
END_PROGRAM

CONFIGURATION Config0
  RESOURCE Res0 ON PLC
    TASK task0(INTERVAL := T#20ms,PRIORITY := 0);
    PROGRAM instance0 WITH task0 : program0;
  END_RESOURCE
END_CONFIGURATION

(* ---- 357-SDT_TO_TOD.ST ---- *)
TYPE oscat_SDT :
	STRUCT
		YEAR : INT;
		MONTH : INT;
		DAY : INT;
		WEEKDAY : INT;
		HOUR : INT;
		MINUTE : INT;
		SECOND : INT;
		MS : INT;
	END_STRUCT;
END_TYPE

FUNCTION _INT_TO_UDINT:UDINT
	VAR_INPUT
		IN :	INT;
	END_VAR

	_INT_TO_UDINT := DINT_TO_UDINT(INT_TO_DINT(IN));
END_FUNCTION

FUNCTION_BLOCK SDT_TO_TOD_Block

	VAR_INPUT
		DTI :	oscat_SDT;
	END_VAR

	VAR_OUTPUT
		SDT_TO_TOD :	UDINT;
	END_VAR

	SDT_TO_TOD := _INT_TO_UDINT(DTI.HOUR) * UDINT#3600000 + _INT_TO_UDINT(DTI.MINUTE) * UDINT#60000 + _INT_TO_UDINT(DTI.SECOND) * UDINT#1000 + _INT_TO_UDINT(DTI.MS);

END_FUNCTION_BLOCK

PROGRAM program0

	VAR
		DTI :	oscat_SDT;
		SDT_TO_TOD :	UDINT;
		func_block : SDT_TO_TOD_Block;
  	END_VAR
	func_block.DTI  :=	DTI;
	func_block();
	SDT_TO_TOD := func_block.SDT_TO_TOD;

END_PROGRAM

CONFIGURATION Config0

	RESOURCE Res0 ON PLC
		TASK task0(INTERVAL := T#20ms,PRIORITY := 0);
		PROGRAM instance0 WITH task0 : program0;
	END_RESOURCE

END_CONFIGURATION

(* ---- 358-CAPITALIZE.ST ---- *)
FUNCTION_BLOCK CAPITALIZE_Block
	VAR_INPUT
		STR :	STRING;
	END_VAR

	VAR_OUTPUT
		CAPITALIZE :	STRING;
	END_VAR

	VAR
		char :	BYTE;
		char2 :	BYTE;
		pos :	INT;
		L :	INT;
		first :	BOOL;
		str_temp :	STRING;
	END_VAR

	CAPITALIZE := str;
	first := TRUE;
	L := LEN(str);
	FOR pos := 1 TO L DO
		char := INT_TO_BYTE(GET_CHAR(str,pos));
		IF first THEN
			char2 := TO_UPPER(char);
			IF char <> char2 THEN
				str_temp := CAPITALIZE;
				CAPITALIZE := REPLACE(str_temp,BYTE_TO_STRING(char2,'%c'),1,pos);
			END_IF;
		END_IF;
		first := char = BYTE#32;
	END_FOR;

END_FUNCTION_BLOCK

PROGRAM program0
  VAR
    LocalVar0 : STRING;
	LocalOUT  : STRING;
	func_block : CAPITALIZE_Block;
  END_VAR
	func_block.CAPITALIZE := LocalVar0;
	func_block();
	LocalOUT := func_block.CAPITALIZE;

END_PROGRAM

CONFIGURATION Config0
  RESOURCE Res0 ON PLC
    TASK task0(INTERVAL := T#20ms,PRIORITY := 0);
    PROGRAM instance0 WITH task0 : program0;
  END_RESOURCE
END_CONFIGURATION

(* ---- 359-SHR_4E.ST ---- *)
FUNCTION_BLOCK SHR_4E_Block

	VAR_INPUT
		SET :	BOOL;
		D0 :	BOOL;
		CLK :	BOOL;
		RST :	BOOL;
	END_VAR

	VAR_OUTPUT
		Q0 :	BOOL;
		Q1 :	BOOL;
		Q2 :	BOOL;
		Q3 :	BOOL;
	END_VAR

	VAR
		trig :	R_TRIG;
	END_VAR

	trig(clk := clk);

	IF set OR rst THEN
		Q0 := NOT RST;
		Q1 := Q0;
		Q2 := Q0;
		Q3 := Q0;
	ELSIF trig.Q THEN
		Q3 := Q2;
		Q2 := Q1;
		Q1 := Q0;
		Q0 := D0;
	END_IF;

END_FUNCTION_BLOCK

PROGRAM program0

	VAR
		SET :	BOOL;
		D0 :	BOOL;
		CLK :	BOOL;
		RST :	BOOL;
		Q0 :	BOOL;
		Q1 :	BOOL;
		Q2 :	BOOL;
		Q3 :	BOOL;
		func_block : SHR_4E_Block;
	END_VAR
	func_block.SET  :=SET;
	func_block.D0  :=D0;
	func_block.CLK  :=CLK;
	func_block.RST  :=RST;
	func_block();
	Q0 := func_block.Q0;
	Q1 := func_block.Q1;
	Q2 := func_block.Q2;
	Q3 := func_block.Q3;

END_PROGRAM

CONFIGURATION Config0
	RESOURCE Res0 ON PLC
		TASK task0(INTERVAL := T#20ms,PRIORITY := 0);
		PROGRAM instance0 WITH task0 : program0;
	END_RESOURCE
END_CONFIGURATION

(* ---- 360-CCOSH.ST ---- *)
TYPE oscat_complex :
  STRUCT
	re : REAL;
	im : REAL;
  END_STRUCT;
END_TYPE

FUNCTION COSH:REAL
	VAR_INPUT
		X :	REAL;
	END_VAR

	VAR
		t :	REAL;
	END_VAR

	T := EXP(X);
	COSH := (1.0 / T + T) * 0.5;
END_FUNCTION

FUNCTION SINH:REAL
	VAR_INPUT
		X :	REAL;
	END_VAR

	IF ABS(x) < 2.0E-3 THEN
		SINH := X;
	ELSE
		SINH := (EXP(x) - EXP(-x)) * 0.5;
	END_IF;
END_FUNCTION

FUNCTION_BLOCK CCOSH_Block
	VAR_INPUT
		X :	oscat_complex;
	END_VAR

	VAR_OUTPUT
		CCOSH :	oscat_complex;
	END_VAR

	CCOSH.re := cosH(x.re) * COS(x.im);
	CCOSH.im := sinH(x.re) * SIN(x.im);
END_FUNCTION_BLOCK

PROGRAM program0
  VAR
    LocalVar0 : oscat_complex;
	LocalOUT  : oscat_complex;
	func_block : CCOSH_Block;
  END_VAR
	func_block.X  := LocalVar0;
	func_block();
	LocalOUT := func_block.CCOSH;
END_PROGRAM

CONFIGURATION Config0
  RESOURCE Res0 ON PLC
    TASK task0(INTERVAL := T#20ms,PRIORITY := 0);
    PROGRAM instance0 WITH task0 : program0;
  END_RESOURCE
END_CONFIGURATION

(* ---- 361-CSINH.ST ---- *)
TYPE oscat_complex :
  STRUCT
	re : REAL;
	im : REAL;
  END_STRUCT;
END_TYPE

FUNCTION COSH:REAL
	VAR_INPUT
		X :	REAL;
	END_VAR

	VAR
		t :	REAL;
	END_VAR

	T := EXP(X);
	COSH := (1.0 / T + T) * 0.5;
END_FUNCTION

FUNCTION SINH:REAL
	VAR_INPUT
		X :	REAL;
	END_VAR

	IF ABS(x) < 2.0E-3 THEN
		SINH := X;
	ELSE
		SINH := (EXP(x) - EXP(-x)) * 0.5;
	END_IF;
END_FUNCTION

FUNCTION_BLOCK CSINH_Block

	VAR_INPUT
		X :	oscat_complex;
	END_VAR

	VAR_OUTPUT
		CSINH :	oscat_complex;
	END_VAR

	CSINH.re := sinH(X.re) * COS(X.im);
	CSINH.im := cosH(X.re) * SIN(X.im);

END_FUNCTION_BLOCK

PROGRAM program0
  VAR
    LocalVar0 : oscat_complex;
	LocalOUT  : oscat_complex;
	func_block : CSINH_Block;
  END_VAR
	func_block.X  := LocalVar0;
	func_block();
	LocalOUT := func_block.CSINH;
END_PROGRAM

CONFIGURATION Config0
  RESOURCE Res0 ON PLC
    TASK task0(INTERVAL := T#20ms,PRIORITY := 0);
    PROGRAM instance0 WITH task0 : program0;
  END_RESOURCE
END_CONFIGURATION

(* ---- 362-MD5_STR.ST ---- *)
FUNCTION_BLOCK MD5_STR

	VAR_INPUT
		RUN :	BOOL;
	END_VAR

	VAR_OUTPUT
		DONE :	BOOL;
	END_VAR

	VAR_IN_OUT
		STR :	oscat_STRING250;
		MD5 :	oscat_aB0_15;
	END_VAR

	VAR
		run_last :	BOOL;
		buf :	oscat_aB0_63;
		mode :	INT;
		size :	UDINT;
		pos :	UDINT;
		i :	INT;
		i2 :	INT;
		MD5_STREAM :	MD5_STREAM;
		CODE :	CODE;
	END_VAR

	CASE mode OF
	0:
		IF RUN AND NOT run_last THEN
			DONE := FALSE;
			mode := 1;
			size := INT_TO_UDINT(LEN(STR));
		END_IF;

	2:
		IF size > UDINT#0 THEN
			i2 := 0;
			FOR i := 1 TO UDINT_TO_INT(SIZE) DO
				CODE(STR:=MID(STR,1,UDINT_TO_INT(POS) + i),POS:=1);
				buf[i2] := CODE.CODE;
				i2 := i2 + 1;
			END_FOR;
		END_IF;

	3:	DONE := TRUE;
		mode := 0;

	END_CASE;

	IF mode > 0 THEN
		MD5_STREAM(SIZE:=size, MODE:=mode, BUF:=buf, MD5:=MD5);
		mode := MD5_STREAM.MODE;
		buf := MD5_STREAM.BUF;
		MD5 := MD5_STREAM.MD5;
		size := MD5_STREAM.SIZE;
		pos := MD5_STREAM.POS;
	END_IF;

	run_last := RUN;

END_FUNCTION_BLOCK

(* ---- 364-CTRL_OUT.ST ---- *)
FUNCTION_BLOCK CTRL_OUT
	VAR_INPUT
		CI :	REAL;
		OFFSET :	REAL;
		MAN_IN :	REAL;
		LIM_L :	REAL;
		LIM_H :	REAL;
		MANUAL :	BOOL;
	END_VAR

	VAR_OUTPUT
		Y :	REAL;
		LIM :	BOOL;
	END_VAR

	Y := SEL(manual, CI, MAN_IN) + OFFSET;

	IF Y >= LIM_H THEN
		Y := LIM_H;
		LIM := TRUE;
	ELSIF Y <= lim_L THEN
		Y := LIM_L;
		LIM := TRUE;
	ELSE
		LIM := FALSE;
	END_IF;
END_FUNCTION_BLOCK

PROGRAM program0
  VAR
	CI :	REAL;
	OFFSET :	REAL;
	MAN_IN :	REAL;
	LIM_L :	REAL;
	LIM_H :	REAL;
	MANUAL :	BOOL;

	Y :	REAL;
	LIM :	BOOL;

	func_block : CTRL_OUT;
  END_VAR
	func_block.CI  := CI ;
	func_block.OFFSET   :=OFFSET ;
	func_block.MAN_IN   :=MAN_IN ;
	func_block.LIM_L   :=LIM_L ;
	func_block.LIM_H   :=LIM_H ;
	func_block.MANUAL   :=MANUAL ;
	func_block();
	Y := func_block.Y;
	LIM := func_block.LIM;
END_PROGRAM

CONFIGURATION Config0
  RESOURCE Res0 ON PLC
    TASK task0(INTERVAL := T#20ms,PRIORITY := 0);
    PROGRAM instance0 WITH task0 : program0;
  END_RESOURCE
END_CONFIGURATION

(* ---- 366-HEX_TO_BYTE.ST ---- *)
TYPE
	 oscat_STRING5  : STRING;
END_TYPE

FUNCTION_BLOCK HEX_TO_BYTE_Block

	VAR_INPUT
		HEX :	oscat_STRING5;
	END_VAR

	VAR_OUTPUT
		HEX_TO_BYTE :	BYTE;
	END_VAR

	VAR
		i :	INT;
		stop :	INT;
		X :	INT;
	END_VAR

	HEX_TO_BYTE := BYTE#0;
	stop := LEN(HEX);
	FOR I := 1 TO stop DO
		x := GET_CHAR(Hex,I);
		IF X > 47 AND x < 58 THEN
			HEX_TO_BYTE := SHL(HEX_TO_BYTE,4) OR INT_TO_BYTE (X - 48);
		ELSIF X > 64 AND X < 71 THEN
			HEX_TO_BYTE := SHL(HEX_TO_BYTE,4) OR INT_TO_BYTE (X - 55);
		ELSIF X > 96 AND X < 103 THEN
			HEX_TO_BYTE := SHL(HEX_TO_BYTE,4) OR INT_TO_BYTE (X - 87);
		END_IF;
	END_FOR;

END_FUNCTION_BLOCK

PROGRAM program0
  VAR
	HEX :	oscat_STRING5;
	HEX_TO_BYTE :	BYTE;
	func_block : HEX_TO_BYTE_Block;
  END_VAR
	func_block.HEX  :=HEX;
	func_block();
	HEX_TO_BYTE := func_block.HEX_TO_BYTE;
END_PROGRAM

CONFIGURATION Config0
	RESOURCE Res0 ON PLC
		TASK task0(INTERVAL := T#20ms,PRIORITY := 0);
		PROGRAM instance0 WITH task0 : program0;
	END_RESOURCE
END_CONFIGURATION

(* ---- 367-ASTRO.ST ---- *)
FUNCTION_BLOCK ASTRO
	VAR_INPUT
		M :	REAL;
		AE :	REAL;
		PC :	REAL;
		LJ :	REAL;
	END_VAR

	VAR_OUTPUT
		YM :	REAL;
		YAE :	REAL;
		YPC :	REAL;
		YLJ :	REAL;
	END_VAR

	YAE :=	AE
			+ m * 6.6845871535E-012
			+ PC * 206265.0
			+ LJ * 63240.0;
	Ym := YAE * 149.597870E9;
	YPC := YAE * 4.8481322570E-006;
	YLJ := YAE * 1.5812776724E-005;
END_FUNCTION_BLOCK

PROGRAM program0
  VAR
    LocalVar0 : REAL;
    LocalVar1 : REAL;
	LocalVar2 : REAL;
	LocalVar3 : REAL;
	LocalOUT1 : REAL;
	LocalOUT2 : REAL;
	LocalOUT3 : REAL;
	LocalOUT4 : REAL;
	func_block : ASTRO;
  END_VAR
	func_block.M  := LocalVar0;
	func_block.AE := LocalVar1;
	func_block.PC := LocalVar2;
	func_block.LJ := LocalVar3;
	func_block();
	LocalOUT1 := func_block.YM ;
	LocalOUT2 := func_block.YAE;
	LocalOUT3 := func_block.YPC;
	LocalOUT4 := func_block.YLJ;

END_PROGRAM

CONFIGURATION Config0
  RESOURCE Res0 ON PLC
    TASK task0(INTERVAL := T#20ms,PRIORITY := 0);
    PROGRAM instance0 WITH task0 : program0;
  END_RESOURCE
END_CONFIGURATION

(* ---- 368-MOON_PHASE.ST ---- *)
FUNCTION TIME_TO_UDINT2:UDINT
	VAR_INPUT
		X :	TIME;
	END_VAR

	TIME_TO_UDINT2 := DINT_TO_UDINT(TIME_TO_DINT(X));
END_FUNCTION

FUNCTION_BLOCK MOON_PHASE_Block

	VAR_INPUT
		XDT :	UDINT;
		SCALE :	BYTE := BYTE#12;
		UPDATE :	TIME := T#1h;
	END_VAR

	VAR_OUTPUT
		PHASE :	BYTE;
	END_VAR

	VAR
		x :	UDINT;
		last_dt :	UDINT;
	END_VAR

	IF XDT - last_dt > TIME_TO_UDINT2(UPDATE) THEN
		x := (XDT - UDINT#603240) MOD UDINT#2551392;
		PHASE := UDINT_TO_BYTE(BYTE_TO_UDINT(SCALE) * x / UDINT#2551392) ;
		last_dt := XDT;
	END_IF;

END_FUNCTION_BLOCK

PROGRAM program0
	VAR
		XDT :	UDINT;
		SCALE :	BYTE := BYTE#12;
		UPDATE :	TIME := T#1h;
		PHASE :	BYTE;

		func_block : MOON_PHASE_Block;
	END_VAR
	func_block.XDT := XDT;
	func_block.SCALE := SCALE;
	func_block.UPDATE := UPDATE;

	func_block();
  	PHASE  := func_block.PHASE;
END_PROGRAM

CONFIGURATION Config0
	RESOURCE Res0 ON PLC
		TASK task0(INTERVAL := T#20ms,PRIORITY := 0);
		PROGRAM instance0 WITH task0 : program0;
	END_RESOURCE
END_CONFIGURATION

(* ---- 369-ARRAY_SPR.ST ---- *)
TYPE
	oscat_pt_ARRAY: ARRAY [1..100] OF REAL;
END_TYPE

FUNCTION_BLOCK ARRAY_SPR_Block
	VAR_IN_OUT
		PT :	oscat_pt_ARRAY;
	END_VAR

	VAR_INPUT
		SIZE :	UINT;
	END_VAR

	VAR_OUTPUT
		ARRAY_SPR :	REAL;
	END_VAR

	VAR
		i :	INT;
		stop :	INT;
		array_max :	REAL;
		array_min :	REAL;
	END_VAR

	stop :=LIMIT_INT(1,UINT_TO_INT(size),1000);

	array_min := pt[1];
	array_max := pt[1];
	FOR i := 2 TO stop DO
		IF pt[i] > array_max THEN array_max := pt[i];
		ELSIF pt[i] < array_min THEN array_min := pt[i];
		END_IF;
	END_FOR;
	array_spr := array_max - array_min;
END_FUNCTION_BLOCK

PROGRAM program0
  VAR
    LocalVar0 : oscat_pt_ARRAY;
    LocalVar1 : UINT;
	LocalOUT  : REAL;
	func_block : ARRAY_SPR_Block;
  END_VAR
	func_block.pt := LocalVar0;
	func_block.size := LocalVar1;
	func_block();
	LocalOUT := func_block.ARRAY_SPR;

END_PROGRAM

CONFIGURATION Config0
  RESOURCE Res0 ON PLC
    TASK task0(INTERVAL := T#20ms,PRIORITY := 0);
    PROGRAM instance0 WITH task0 : program0;
  END_RESOURCE
END_CONFIGURATION

(* ---- 372-ARRAY_VAR.ST ---- *)
TYPE
	oscat_pt_ARRAY: ARRAY [1..100] OF REAL;
END_TYPE

FUNCTION_BLOCK ARRAY_VAR_Block
	VAR_IN_OUT
		PT :	oscat_pt_ARRAY;
	END_VAR

	VAR_INPUT
		SIZE :	UINT;
	END_VAR

	VAR_OUTPUT
		ARRAY_VAR :	REAL;
	END_VAR

	VAR
		i :	INT;
		stop :	INT;
		avg :	REAL;
	END_VAR

	stop :=LIMIT_INT(1,UINT_TO_INT(size),1000);
	avg := pt[1];
	FOR i := 2 TO stop DO
		avg := avg + pt[i];
	END_FOR;
	avg := avg / INT_TO_REAL(stop);

	array_var := EXPT(pt[1] - avg, 2.0);
	FOR i := 2 TO stop DO
		array_var := array_var + EXPT(pt[i] - avg, 2.0);
	END_FOR;
	array_var := array_var / INT_TO_REAL(stop-1);

END_FUNCTION_BLOCK

PROGRAM program0
  VAR
    LocalVar0 : oscat_pt_ARRAY;
    LocalVar1 : UINT;
	LocalOUT  : REAL;
	func_block : ARRAY_VAR_Block;
  END_VAR
	func_block.pt := LocalVar0;
	func_block.size := LocalVar1;
	func_block();
	LocalOUT := func_block.ARRAY_VAR;

END_PROGRAM

CONFIGURATION Config0
  RESOURCE Res0 ON PLC
    TASK task0(INTERVAL := T#20ms,PRIORITY := 0);
    PROGRAM instance0 WITH task0 : program0;
  END_RESOURCE
END_CONFIGURATION

(* ---- 373-CSQRT.ST ---- *)
TYPE oscat_complex :
  STRUCT
	re : REAL;
	im : REAL;
  END_STRUCT;
END_TYPE

FUNCTION HYPOT:REAL
	VAR_INPUT
		X :	REAL;
		Y :	REAL;
	END_VAR

	HYPOT := SQRT(x*x + y*y);
END_FUNCTION

FUNCTION SGN : INT
  VAR_INPUT
    x : REAL;
  END_VAR

  IF X > 0.0 THEN
  	sgn := 1;
  ELSIF X < 0.0 THEN
  	sgn := -1;
  ELSE
  	sgn := 0;
  END_IF;
END_FUNCTION

FUNCTION_BLOCK CSQRT_Block
	VAR_INPUT
		X :	oscat_complex;
	END_VAR

	VAR_OUTPUT
		CSQRT :	oscat_complex;
	END_VAR

	VAR
		temp :	REAL;
	END_VAR

	temp := HYPOT(x.re, x.im);
	CSQRT.re :=  SQRT(0.5 * (temp + x.re));
	CSQRT.im :=  INT_TO_REAL(sgn(x.im)) * SQRT(0.5 * (temp - x.re));

END_FUNCTION_BLOCK

PROGRAM program0
  VAR
    LocalVar0 : oscat_complex;
	LocalOUT  : oscat_complex;
	func_block : CSQRT_Block;
  END_VAR
	func_block.X  := LocalVar0;
	func_block();
	LocalOUT := func_block.CSQRT;
END_PROGRAM

CONFIGURATION Config0
  RESOURCE Res0 ON PLC
    TASK task0(INTERVAL := T#20ms,PRIORITY := 0);
    PROGRAM instance0 WITH task0 : program0;
  END_RESOURCE
END_CONFIGURATION

(* ---- 374-ELEMENT_COUNT.ST ---- *)
TYPE
	oscat_STRING250             : STRING;
END_TYPE

FUNCTION_BLOCK ELEMENT_COUNT_Block

	VAR_IN_OUT
		ELEMENT :	oscat_STRING250;
	END_VAR

	VAR_INPUT
		SEP :	BYTE;
	END_VAR

	VAR_OUTPUT
		ELEMENT_COUNT :	INT;
	END_VAR

	VAR
		I :	INT;
		pos :	INT;
	END_VAR

	i := LEN(ELEMENT);
	IF i = 0 THEN
		ELEMENT_COUNT := 0;
	ELSE
		ELEMENT_COUNT := 1;
		FOR pos := 1 TO I DO
			IF INT_TO_BYTE(GET_CHAR(ELEMENT,pos)) = SEP THEN ELEMENT_COUNT := ELEMENT_COUNT + 1; END_IF;
		END_FOR;
	END_IF;

END_FUNCTION_BLOCK

PROGRAM program0
	VAR
		SEP :	BYTE;
		POS :	INT;
		ELEMENT :	oscat_STRING250;
		ELEMENT_GET :	oscat_STRING250;

		func_block : ELEMENT_COUNT_Block;
	END_VAR
	func_block.SEP    :=SEP    ;
	func_block.POS:=POS;
	func_block.ELEMENT     :=ELEMENT     ;
	func_block();
	ELEMENT    := func_block.ELEMENT    ;
	ELEMENT_GET:= func_block.ELEMENT_GET;

END_PROGRAM

CONFIGURATION Config0
  RESOURCE Res0 ON PLC
    TASK task0(INTERVAL := T#20ms,PRIORITY := 0);
    PROGRAM instance0 WITH task0 : program0;
  END_RESOURCE
END_CONFIGURATION

(* ---- 375-FF_D4E.ST ---- *)
FUNCTION_BLOCK FF_D4E
	VAR_INPUT
		D0 :	BOOL;
		D1 :	BOOL;
		D2 :	BOOL;
		D3 :	BOOL;
		CLK :	BOOL;
		RST :	BOOL;
	END_VAR

	VAR_OUTPUT
		Q0 :	BOOL;
		Q1 :	BOOL;
		Q2 :	BOOL;
		Q3 :	BOOL;
	END_VAR

	VAR
		edge :	BOOL;
	END_VAR

	IF rst THEN
		Q0 := FALSE;
		Q1 := FALSE;
		Q2 := FALSE;
		Q3 := FALSE;
	ELSIF clk AND NOT edge THEN
		Q0 := D0;
		Q1 := D1;
		Q2 := D2;
		Q3 := D3;
	END_IF;
	edge := CLK;
END_FUNCTION_BLOCK

PROGRAM program0
  VAR
		D0  :	BOOL;
		D1  :	BOOL;
		D2  :	BOOL;
		D3  :	BOOL;
		CLK :	BOOL;
		RST :	BOOL;

		Q0 :	BOOL;
		Q1 :	BOOL;
		Q2 :	BOOL;
		Q3 :	BOOL;

	func_block : FF_D4E;
  END_VAR
	func_block.D0 :=D0 ;
	func_block.D1 :=D1 ;
	func_block.D2 :=D2 ;
	func_block.D3 :=D3 ;
	func_block.CLK:=CLK;
	func_block.RST:=RST;
	func_block();
	Q0 := func_block.Q0;
	Q1 := func_block.Q1;
	Q2 := func_block.Q2;
	Q3 := func_block.Q3;
END_PROGRAM

CONFIGURATION Config0
  RESOURCE Res0 ON PLC
    TASK task0(INTERVAL := T#20ms,PRIORITY := 0);
    PROGRAM instance0 WITH task0 : program0;
  END_RESOURCE
END_CONFIGURATION

(* ---- 376-CARG.ST ---- *)
TYPE oscat_complex :
  STRUCT
	re : REAL;
	im : REAL;
  END_STRUCT;
END_TYPE

FUNCTION ATAN2:REAL
	VAR_INPUT
		X :	REAL;
		Y :	REAL;
	END_VAR

	IF X > 0.0 THEN
		ATAN2 := ATAN(Y/X);
	ELSIF X < 0.0 THEN
		IF Y >= 0.0 THEN
			ATAN2 := ATAN(Y/X) + 3.14159265358979323846264338327950288;
		ELSE
			ATAN2 := ATAN(Y/X) - 3.14159265358979323846264338327950288;
		END_IF;
	ELSIF Y > 0.0 THEN
		ATAN2 := 1.5707963267948965580;
	ELSIF Y < 0.0 THEN
		ATAN2 := -1.5707963267948965580;
	ELSE
		ATAN2 := 0.0;
	END_IF;

END_FUNCTION

FUNCTION_BLOCK CARG_Block

	VAR_INPUT
		X :	oscat_complex;
	END_VAR

	VAR_OUTPUT
		CARG :	REAL;
	END_VAR

	CARG := ATAN2(X.im, X.re);

END_FUNCTION_BLOCK

PROGRAM program0
  VAR
    LocalVar0 : oscat_complex;
	LocalOUT  : REAL;
	func_block : CARG_Block;
  END_VAR
	func_block.X  := LocalVar0;
	func_block();
	LocalOUT := func_block.CARG;
END_PROGRAM

CONFIGURATION Config0
  RESOURCE Res0 ON PLC
    TASK task0(INTERVAL := T#20ms,PRIORITY := 0);
    PROGRAM instance0 WITH task0 : program0;
  END_RESOURCE
END_CONFIGURATION

(* ---- 377-INSERT250.ST ---- *)
TYPE
	oscat_STRING250             : STRING;
END_TYPE

FUNCTION_BLOCK _INSERT250
    VAR_INPUT
        IN1 :	oscat_STRING250;
        IN2 :	oscat_STRING250;
        P :	INT;
    END_VAR
    VAR_OUTPUT
        _INSERT :	oscat_STRING250;
    END_VAR
    VAR
        size :	INT;
    END_VAR

    size := LEN(IN1);
    IF size + LEN(IN2) <= 250 THEN
        P := LIMIT(0,P,size);
        IF P = 0 THEN
            _INSERT := CONCAT(IN2,IN1);
        ELSE
            _INSERT := INSERT(IN1, IN2, P);
        END_IF;
    END_IF;

END_FUNCTION_BLOCK

PROGRAM program0
	VAR
	    LocalVar1 : oscat_STRING250;
        LocalVar2 : oscat_STRING250;
        LocalVar3 : INT;
		LocalOUT  : oscat_STRING250;
		func_block : _INSERT250;
  	END_VAR
	func_block.IN1 := LocalVar1;
    func_block.IN2 := LocalVar2;
    func_block.P := LocalVar3;
	func_block();
	LocalOUT := func_block._INSERT;
END_PROGRAM

CONFIGURATION Config0
  	RESOURCE Res0 ON PLC
    	TASK task0(INTERVAL := T#20ms,PRIORITY := 0);
    	PROGRAM instance0 WITH task0 : program0;
  	END_RESOURCE
END_CONFIGURATION

(* ---- 378-LINEAR_INT.ST ---- *)
TYPE
	oscat_ARRAY_X               : ARRAY [0..1]    OF REAL;
	oscat_XY                    : ARRAY [1..20]   OF oscat_ARRAY_X := [0,0,0,0,0,0,0,0,0,0,0,0,0,0,0,0,0,0,0,0];
END_TYPE

FUNCTION_BLOCK LINEAR_INT_Block

	VAR_INPUT
		X :	REAL;
		XY :	oscat_XY;
		PTS :	INT;
	END_VAR

	VAR_OUTPUT
		LINEAR_INT :	REAL;
	END_VAR

	VAR
		i :	INT;
		i2 :	INT;
	END_VAR

	pts := MIN(pts,20);

	i := 2;

	WHILE (i < pts) AND (XY[i][0] < X) DO
		i := i + 1;
	END_WHILE;

	i2 := i-1;

	LINEAR_INT := ((XY[i][1] - XY[i2][1]) * X - XY[i][1] * XY[i2][0] + XY[i2][1] * XY[i][0]) / (XY[i][0] - XY[i2][0]);

END_FUNCTION_BLOCK

PROGRAM program0

	VAR
		X :	REAL;
		XY :	oscat_XY;
		PTS :	INT;

		LINEAR_INT :	REAL;

		func_block : LINEAR_INT_Block;
	END_VAR
	func_block.X := X;
	func_block.XY := XY;
	func_block.PTS := PTS;

	func_block();
	LINEAR_INT := func_block.LINEAR_INT;

END_PROGRAM

CONFIGURATION Config0

	RESOURCE Res0 ON PLC
		TASK task0(INTERVAL := T#20ms,PRIORITY := 0);
		PROGRAM instance0 WITH task0 : program0;
	END_RESOURCE

END_CONFIGURATION

(* ---- 379-MANUAL_2.ST ---- *)
FUNCTION_BLOCK MANUAL_2_Block

	VAR_INPUT
		_IN :	BOOL;
		ENA :	BOOL;
		_ON :	BOOL;
		OFF :	BOOL;
		MAN :	BOOL;
	END_VAR

	VAR_OUTPUT
		Q :	BOOL;
		STATUS :	BYTE;
	END_VAR

	IF ena THEN
		IF NOT _ON AND NOT OFF THEN
			Q := _IN;
			STATUS := BYTE#100;
		ELSIF _on AND NOT off THEN
			Q := TRUE;
			STATUS := BYTE#101;
		ELSIF NOT _on AND off THEN
			q := FALSE;
			STATUS := BYTE#102;
		ELSE
			Q := MAN;
			STATUS := BYTE#103;
		END_IF;
	ELSE
		Q := FALSE;
		STATUS := BYTE#104;
	END_IF;

END_FUNCTION_BLOCK

PROGRAM program0

	VAR
		_IN :	BOOL;
		ENA :	BOOL;
		_ON :	BOOL;
		OFF :	BOOL;
		MAN :	BOOL;

		Q :	BOOL;
		STATUS :	BYTE;

		func_block : MANUAL_2_Block;
	END_VAR
	func_block._IN := _IN;
	func_block.ENA := ENA;
	func_block._ON := _ON;
	func_block.OFF := OFF;
	func_block.MAN := MAN;
	func_block();
	Q := func_block.Q;
	STATUS := func_block.STATUS;

END_PROGRAM

CONFIGURATION Config0

	RESOURCE Res0 ON PLC
		TASK task0(INTERVAL := T#20ms,PRIORITY := 0);
		PROGRAM instance0 WITH task0 : program0;
	END_RESOURCE

END_CONFIGURATION

(* ---- 380-LTCH_4.ST ---- *)
FUNCTION_BLOCK LTCH_4_Block

	VAR_INPUT
		D0 :	BOOL;
		D1 :	BOOL;
		D2 :	BOOL;
		D3 :	BOOL;
		L :	BOOL;
		RST :	BOOL;
	END_VAR

	VAR_OUTPUT
		Q0 :	BOOL;
		Q1 :	BOOL;
		Q2 :	BOOL;
		Q3 :	BOOL;
	END_VAR

	IF rst THEN			(* if asynchronous reset then Q=0 *)
		Q0 := FALSE;
		Q1 := FALSE;
		Q2 := FALSE;
		Q3 := FALSE;
	ELSIF L THEN			(* latch is transparent *)
		Q0 := D0;
		Q1 := D1;
		Q2 := D2;
		Q3 := D3;
	END_IF;

END_FUNCTION_BLOCK

PROGRAM program0

	VAR
		D0 :	BOOL;
		D1 :	BOOL;
		D2 :	BOOL;
		D3 :	BOOL;
		L :	BOOL;
		RST :	BOOL;

		Q0 :	BOOL;
		Q1 :	BOOL;
		Q2 :	BOOL;
		Q3 :	BOOL;

		func_block : LTCH_4_Block;
	END_VAR
	func_block.D0 := D0;
	func_block.D1 := D1;
	func_block.D2 := D2;
	func_block.D3 := D3;
	func_block.L := L;
	func_block.RST := RST;

	func_block();
	Q0 := func_block.Q0;
	Q1 := func_block.Q1;
	Q2 := func_block.Q2;
	Q3 := func_block.Q3;

END_PROGRAM

CONFIGURATION Config0

	RESOURCE Res0 ON PLC
		TASK task0(INTERVAL := T#20ms,PRIORITY := 0);
		PROGRAM instance0 WITH task0 : program0;
	END_RESOURCE

END_CONFIGURATION

(* ---- 381-DRIVER_1.ST ---- *)
FUNCTION_BLOCK DRIVER_1
	VAR_INPUT
		SET :	BOOL;
		IN :	BOOL;
		RST :	BOOL;
		TOGGLE_MODE :	BOOL;
		TIMEOUT :	TIME;
	END_VAR

	VAR_OUTPUT
		Q :	BOOL;
	END_VAR

	VAR
		off :	TON;
		edge :	BOOL;
	END_VAR

	IF off.Q THEN Q := FALSE; END_IF;
	IF rst THEN
		Q := FALSE;
	ELSIF set THEN
		Q := TRUE;
	ELSIF IN AND NOT edge THEN
		IF toggle_mode THEN q := NOT Q; ELSE q := TRUE; END_IF;
	END_IF;
	edge := in;
	IF timeout > t#0s THEN off(in := Q, PT := Timeout); END_IF;

END_FUNCTION_BLOCK

PROGRAM program0
  VAR
	SET         :	BOOL;
	IN          :	BOOL;
	RST         :	BOOL;
	TOGGLE_MODE :	BOOL;
	TIMEOUT     :	TIME;

	Q :	BOOL;

	func_block : DRIVER_1;
  END_VAR
	func_block.SET         :=SET        ;
	func_block.IN          :=IN         ;
	func_block.RST         :=RST        ;
	func_block.TOGGLE_MODE :=TOGGLE_MODE;
	func_block.TIMEOUT     :=TIMEOUT    ;
	func_block();
	Q := func_block.Q;
END_PROGRAM

CONFIGURATION Config0
  RESOURCE Res0 ON PLC
    TASK task0(INTERVAL := T#20ms,PRIORITY := 0);
    PROGRAM instance0 WITH task0 : program0;
  END_RESOURCE
END_CONFIGURATION

(* ---- 382-DELAY.ST ---- *)
TYPE
	oscat_delay_buf             : ARRAY [0..31]   OF REAL;
END_TYPE

FUNCTION INC1:INT

	VAR_INPUT
		X :	INT;
		N :	INT;
	END_VAR

	IF X >= N - 1 THEN
		INC1 := 0;
	ELSE
		INC1 := X + 1;
	END_IF;
END_FUNCTION

FUNCTION_BLOCK DELAY

	VAR_INPUT
		IN :	REAL;
		N :	INT;
		RST :	BOOL;
	END_VAR

	VAR_OUTPUT
		OUT :	REAL;
	END_VAR

	VAR
		buf :	oscat_delay_buf;
		i :	INT;
		init :	BOOL;
		stop :	INT;
	END_VAR

	stop := LIMIT(0,N,32) - 1;
	IF rst OR NOT init THEN
		init := TRUE;
		FOR i := 0 TO stop DO buf[i] := in; END_FOR;
		out := in;
		i := 0;
	ELSIF stop < 0 THEN
		out := in;
	ELSE
		out := buf[i];
		buf[i] := in;
		i := INC1(i, N);
	END_IF;

END_FUNCTION_BLOCK

PROGRAM program0
  VAR
	IN :	REAL;
	N :	INT;
	RST :	BOOL;
	OUT :	REAL;
	func_block : DELAY;
  END_VAR
	func_block.IN  :=IN;
	func_block.N  :=N;
	func_block.RST  :=RST;
	func_block();
	OUT := func_block.OUT;

END_PROGRAM

CONFIGURATION Config0
	RESOURCE Res0 ON PLC
		TASK task0(INTERVAL := T#20ms,PRIORITY := 0);
		PROGRAM instance0 WITH task0 : program0;
	END_RESOURCE
END_CONFIGURATION

(* ---- 383-INC_DEC.ST ---- *)
FUNCTION_BLOCK INC_DEC_Block

	VAR_INPUT
		CHA :	BOOL;
		CHB :	BOOL;
		RST :	BOOL := 0;
	END_VAR

	VAR_OUTPUT
		DIR :	BOOL;
		CNT :	INT;
	END_VAR

	VAR
		edgea :	BOOL := 0;
		clk :	BOOL;
		clka :	BOOL;
		clkb :	BOOL;
		edgeb :	BOOL;
		axb :	BOOL;
	END_VAR

	axb := cha XOR chb;

	clka := cha XOR edgea;
	edgea := cha;

	clkb := chb XOR edgeb;
	edgeb := chb;

	clk := clka OR clkb;

	IF axb AND clka THEN dir := TRUE; END_IF;
	IF axb AND clkb THEN dir := FALSE; END_IF;

	IF clk AND dir THEN cnt := cnt + 1; END_IF;
	IF clk AND NOT dir THEN cnt := cnt -1; END_IF;

	IF rst THEN cnt := 0; END_IF;

END_FUNCTION_BLOCK

PROGRAM program0

	VAR
		CHA :	BOOL;
		CHB :	BOOL;
		RST :	BOOL := 0;

		DIR :	BOOL;
		CNT :	INT;
		func_block : INC_DEC_Block;
	END_VAR
	func_block.CHA := CHA;
	func_block.CHB := CHB;
	func_block.RST := RST;
	func_block();
	DIR := func_block.DIR;
	CNT := func_block.CNT;

END_PROGRAM

CONFIGURATION Config0

	RESOURCE Res0 ON PLC
		TASK task0(INTERVAL := T#20ms,PRIORITY := 0);
		PROGRAM instance0 WITH task0 : program0;
	END_RESOURCE

END_CONFIGURATION

(* ---- 386-CTAN.ST ---- *)
TYPE oscat_complex :
  STRUCT
	re : REAL;
	im : REAL;
  END_STRUCT;
END_TYPE

FUNCTION COSH:REAL
	VAR_INPUT
		X :	REAL;
	END_VAR

	VAR
		t :	REAL;
	END_VAR

	T := EXP(X);
	COSH := (1.0 / T + T) * 0.5;
END_FUNCTION

FUNCTION SINH:REAL
	VAR_INPUT
		X :	REAL;
	END_VAR

	IF ABS(x) < 2.0E-3 THEN
		SINH := X;
	ELSE
		SINH := (EXP(x) - EXP(-x)) * 0.5;
	END_IF;
END_FUNCTION

FUNCTION_BLOCK CTAN_Block
	VAR_INPUT
		X :	oscat_complex;
	END_VAR

	VAR_OUTPUT
		CTAN :	oscat_complex;
	END_VAR

	VAR
		temp :	REAL;
		xi2 :	REAL;
		xr2 :	REAL;
	END_VAR

	xi2 := 2.0 * x.im;
	xr2 := 2.0 * x.re;
	temp := 1.0 / (COS(xr2) + COSH( xi2));
	CTAN.re := temp * SIN(xr2);
	CTAN.im := temp * SINH(xi2);
END_FUNCTION_BLOCK

PROGRAM program0
  VAR
    LocalVar0 : oscat_complex;
	LocalOUT  : oscat_complex;
	func_block : CTAN_Block;
  END_VAR
	func_block.X  := LocalVar0;
	func_block();
	LocalOUT := func_block.CTAN;
END_PROGRAM

CONFIGURATION Config0
  RESOURCE Res0 ON PLC
    TASK task0(INTERVAL := T#20ms,PRIORITY := 0);
    PROGRAM instance0 WITH task0 : program0;
  END_RESOURCE
END_CONFIGURATION

(* ---- 387-TEMPERATURE.ST ---- *)
FUNCTION_BLOCK TEMPERATURE

	VAR_INPUT
		K :	REAL;
		C :	REAL := -273.15;
		F :	REAL := -459.67;
		RE :	REAL := -218.52;
		RA :	REAL := 0.0;
	END_VAR

	VAR_OUTPUT
		YK :	REAL;
		YC :	REAL;
		YF :	REAL;
		YRE :	REAL;
		YRA :	REAL;
	END_VAR

	YK := K + (C + 273.15) + (F + 459.67) * 0.555555555555 + (Re * 1.25 + 273.15) + (Ra * 0.555555555555);
	YC := YK -273.15;
	YF := YK * 1.8 - 459.67;
	YRe := (YK - 273.15) * 0.8;
	YRa := YK * 1.8;

END_FUNCTION_BLOCK

PROGRAM program0
  VAR
	K :	REAL;
	C :	REAL := -273.15;
	F :	REAL := -459.67;
	RE :	REAL := -218.52;
	RA :	REAL := 0.0;
	YK :	REAL;
	YC :	REAL;
	YF :	REAL;
	YRE :	REAL;
	YRA :	REAL;
	func_block : TEMPERATURE;
  END_VAR
	func_block.K  :=K;
	func_block.C  :=C;
	func_block.F  :=F;
	func_block.RE  :=RE;
	func_block.RA  :=RA;
	func_block();
	YK := func_block.YK;
	YC := func_block.YC;
	YF := func_block.YF;
	YRE := func_block.YRE;
	YRA := func_block.YRA;

END_PROGRAM

CONFIGURATION Config0
	RESOURCE Res0 ON PLC
		TASK task0(INTERVAL := T#20ms,PRIORITY := 0);
		PROGRAM instance0 WITH task0 : program0;
	END_RESOURCE
END_CONFIGURATION

(* ---- 388-REPLACE_CHARS.ST ---- *)
FUNCTION_BLOCK REPLACE_CHARS_Block

	VAR_INPUT
		STR :	STRING;
		SRC :	STRING;
		REP :	STRING;
	END_VAR

	VAR_OUTPUT
		REPLACE_CHARS :	STRING;
	END_VAR

	VAR
		tmp :	STRING;
		a :	INT;
		b :	INT;
		c :	STRING;
		stp :	INT;
	END_VAR

	REPLACE_CHARS := STR;

	a := LEN(src);
	b := LEN(rep);
	IF a < b THEN
		rep := LEFT(rep, a);
	ELSIF b < a THEN
		src := LEFT(src, b);
	END_IF;

	stp := LEN(str);
	FOR a := 1 TO stp DO
		c := MID(REPLACE_CHARS, 1, a);
		b := FIND(src, c);
		IF b > 0 THEN
			tmp := MID(rep, 1, b);
			REPLACE_CHARS := REPLACE(REPLACE_CHARS, tmp, 1, a);
		END_IF;
	END_FOR;

END_FUNCTION_BLOCK

PROGRAM program0

	VAR
		STR :	STRING;
		SRC :	STRING;
		REP :	STRING;

        REPLACE_CHARS :	STRING;
		func_block : REPLACE_CHARS_Block;
	END_VAR
		func_block.STR := STR;
		func_block.SRC := SRC;
		func_block.REP := REP;
		func_block();
		REPLACE_CHARS := func_block.REPLACE_CHARS;

END_PROGRAM

CONFIGURATION Config0

	RESOURCE Res0 ON PLC
		TASK task0(INTERVAL := T#20ms,PRIORITY := 0);
		PROGRAM instance0 WITH task0 : program0;
	END_RESOURCE

END_CONFIGURATION

(* ---- 389-CTANH.ST ---- *)
TYPE oscat_complex :
  STRUCT
	re : REAL;
	im : REAL;
  END_STRUCT;
END_TYPE

FUNCTION COSH:REAL
	VAR_INPUT
		X :	REAL;
	END_VAR

	VAR
		t :	REAL;
	END_VAR

	T := EXP(X);
	COSH := (1.0 / T + T) * 0.5;
END_FUNCTION

FUNCTION SINH:REAL
	VAR_INPUT
		X :	REAL;
	END_VAR

	IF ABS(x) < 2.0E-3 THEN
		SINH := X;
	ELSE
		SINH := (EXP(x) - EXP(-x)) * 0.5;
	END_IF;
END_FUNCTION

FUNCTION_BLOCK CTANH_Block
	VAR_INPUT
		X :	oscat_complex;
	END_VAR

	VAR_OUTPUT
		CTANH :	oscat_complex;
	END_VAR

	VAR
		xi2 :	REAL;
		xr2 :	REAL;
		temp :	REAL;
	END_VAR

	xi2 := 2.0 * x.im;
	xr2 := 2.0 * x.re;
	temp := 1.0 /(COSH(xr2) + COS(xi2));
	CTANH.re := temp * SINH(xr2);
	CTANH.im := temp * SIN(xi2);

END_FUNCTION_BLOCK

PROGRAM program0
  VAR
    LocalVar0 : oscat_complex;
	LocalOUT  : oscat_complex;
	func_block : CTANH_Block;
  END_VAR
	func_block.X  := LocalVar0;
	func_block();
	LocalOUT := func_block.CTANH;
END_PROGRAM

CONFIGURATION Config0
  RESOURCE Res0 ON PLC
    TASK task0(INTERVAL := T#20ms,PRIORITY := 0);
    PROGRAM instance0 WITH task0 : program0;
  END_RESOURCE
END_CONFIGURATION

(* ---- 390-LIST_ADD.ST ---- *)
FUNCTION_BLOCK CHR_TO_STRING_Block
	VAR_INPUT
		C :	BYTE;
	END_VAR

	VAR_OUTPUT
		CHR_TO_STRING :	STRING;
	END_VAR

	CHR_TO_STRING := BYTE_TO_STRING(C);

END_FUNCTION_BLOCK

FUNCTION_BLOCK LIST_ADD_Block

	VAR_INPUT
		SEP :	BYTE;
		INS :	STRING;
	END_VAR

	VAR_IN_OUT
		LIST :	STRING;
	END_VAR

	VAR_OUTPUT
		LIST_ADD :	BOOL;
	END_VAR

	VAR
		CHR_TO_STRING :	CHR_TO_STRING_Block;
	END_VAR

	IF LEN(LIST) + LEN(INS) + 1 <= 250 THEN
	CHR_TO_STRING(C:=SEP);
	LIST := CONCAT(LIST, CHR_TO_STRING.CHR_TO_STRING);
	LIST := CONCAT(LIST, INS);
	LIST_ADD := TRUE;
	ELSE
	LIST_ADD := FALSE;
	END_IF;

END_FUNCTION_BLOCK

PROGRAM program0

	VAR
		SEP :	BYTE;
		INS :	STRING;

		LIST :	STRING;

		LIST_ADD :	BOOL;

		func_block : LIST_ADD_Block;
	END_VAR
	func_block.SEP := SEP;
	func_block.INS := INS;
	func_block.LIST := LIST;

	func_block();
	LIST := func_block.LIST;
	LIST_ADD := func_block.LIST_ADD;

END_PROGRAM

CONFIGURATION Config0

	RESOURCE Res0 ON PLC
		TASK task0(INTERVAL := T#20ms,PRIORITY := 0);
		PROGRAM instance0 WITH task0 : program0;
	END_RESOURCE

END_CONFIGURATION

(* ---- 391-IP4_DECODE.ST ---- *)
TYPE
  oscat_STRING80             : STRING;
END_TYPE

FUNCTION_BLOCK IP4_DECODE_Block

	VAR_INPUT
		STR :	oscat_STRING80;
	END_VAR

	VAR_OUTPUT
		IP4_DECODE :	DWORD;
	END_VAR

	VAR
		pos :	INT;
		IS_NUM :	IS_NUM;
	END_VAR

	IP4_DECODE := DWORD#0;
	pos := FIND(str, '.');
	WHILE pos > 0 DO
		IP4_DECODE := SHL(IP4_DECODE,8);
		IF POS > 1 AND POS <= 4 THEN
			IS_NUM(STR:=LEFT(str,pos - 1));
			IF IS_NUM.IS_NUM THEN
				IP4_DECODE := IP4_DECODE OR STRING_TO_DWORD(IS_NUM.STR);
			END_IF;
		END_IF;
		str := DELETE(str, pos, 1);
		pos := FIND(str, '.');
	END_WHILE;

	IP4_DECODE := SHL(IP4_DECODE,8);
	IS_NUM(STR:=str);
	IF IS_NUM.IS_NUM THEN
	IP4_DECODE := IP4_DECODE OR STRING_TO_DWORD(str);
	END_IF;

END_FUNCTION_BLOCK

PROGRAM program0
	VAR
		STR :	oscat_STRING80;
		IP4_DECODE :	DWORD;

		func_block : IP4_DECODE_Block;
	END_VAR
	func_block.STR := STR;

	func_block();
	IP4_DECODE  := func_block.IP4_DECODE;
END_PROGRAM

CONFIGURATION Config0

  	RESOURCE Res0 ON PLC
    	TASK task0(INTERVAL := T#20ms,PRIORITY := 0);
    	PROGRAM instance0 WITH task0 : program0;
  	END_RESOURCE

END_CONFIGURATION

(* ---- 392-ARRAY_GAV.ST ---- *)
TYPE
	oscat_pt_ARRAY: ARRAY [1..100] OF REAL;
END_TYPE

FUNCTION SQRTN:REAL
	VAR_INPUT
		X :	REAL;
		N :	INT;
	END_VAR

	IF N > 0 THEN
		SQRTN := EXP(LN(x) / INT_TO_REAL(n));
	ELSE
		SQRTN := 0.0;
	END_IF;
END_FUNCTION

FUNCTION_BLOCK ARRAY_GAV_Block
	VAR_IN_OUT
		PT :	oscat_pt_ARRAY;
	END_VAR

	VAR_INPUT
		SIZE :	UINT;
	END_VAR

	VAR_OUTPUT
		ARRAY_GAV :	REAL;
	END_VAR

	VAR
		i :	INT;
		stop :	INT;
	END_VAR

	stop :=LIMIT_INT(1,UINT_TO_INT(size),1000);
	ARRAY_GAV := 1.0;
	FOR i := 1 TO stop DO
		IF pt[i] > 0.0 THEN
			ARRAY_GAV := ARRAY_GAV * pt[i];
		ELSE
			ARRAY_GAV := 0.0;
			RETURN;
		END_IF;
	END_FOR;
	ARRAY_GAV := SQRTN(ARRAY_GAV,stop);
END_FUNCTION_BLOCK

PROGRAM program0
  VAR
    LocalVar0 : oscat_pt_ARRAY;
    LocalVar1 : UINT;
	LocalOUT  : REAL;
	func_block : ARRAY_GAV_Block;
  END_VAR
	func_block.pt := LocalVar0;
	func_block.size := LocalVar1;
	func_block();
	LocalOUT := func_block.ARRAY_GAV;

END_PROGRAM

CONFIGURATION Config0
  RESOURCE Res0 ON PLC
    TASK task0(INTERVAL := T#20ms,PRIORITY := 0);
    PROGRAM instance0 WITH task0 : program0;
  END_RESOURCE
END_CONFIGURATION

(* ---- 393-CLICK_DEC.ST ---- *)
FUNCTION_BLOCK CLICK_DEC

	VAR_INPUT
		IN :	BOOL;
		TC :	TIME;
	END_VAR

	VAR_OUTPUT
		Q0 :	BOOL;
		Q1 :	BOOL;
		Q2 :	BOOL;
		Q3 :	BOOL;
	END_VAR

	VAR
		tx :	TP;
		edge :	BOOL;
		cnt :	INT := INT#-1;
	END_VAR

	IF in = FALSE THEN
		Q0 := FALSE;
		Q1 := FALSE;
		Q2 := FALSE;
		Q3 := FALSE;
	END_IF;

	IF in AND NOT edge AND NOT tx.q THEN
		cnt := 0;
	ELSIF tx.Q AND NOT IN AND edge THEN
		cnt := cnt + 1;
	ELSIF NOT tx.Q THEN
		CASE cnt OF
			0 : Q0 := TRUE;
			1 : Q1 := TRUE;
			2 : Q2 := TRUE;
			3 : Q3 := TRUE;
		END_CASE;
		cnt := -1;
	END_IF;

	edge := IN;
	tx(in := IN, pt := TC);

END_FUNCTION_BLOCK

PROGRAM program0
  VAR
    LocalVar0 : BOOL;
    LocalVar1 : TIME;
	Q0 :	BOOL;
	Q1 :	BOOL;
	Q2 :	BOOL;
	Q3 :	BOOL;
	func_block : CLICK_DEC;
  END_VAR
	func_block.IN  := LocalVar0;
	func_block.TC := LocalVar1;
	func_block();
	Q0 := func_block.Q0;
	Q1 := func_block.Q1;
	Q2 := func_block.Q2;
	Q3 := func_block.Q3;
END_PROGRAM

CONFIGURATION Config0
  RESOURCE Res0 ON PLC
    TASK task0(INTERVAL := T#20ms,PRIORITY := 0);
    PROGRAM instance0 WITH task0 : program0;
  END_RESOURCE
END_CONFIGURATION
